METHOD PRIVATE Test_EStopRequestSwitchesOutputsOffAndBlocksRestart
TcUnit.TEST(__POUNAME());
// arrange: running
group_3(Run := TRUE);
fb_3(Restart := FALSE, EStopIn1 := TRUE, EStopIn2 := TRUE);
group_3(Run := TRUE);
fb_3(Restart := TRUE, EStopIn1 := TRUE, EStopIn2 := TRUE);
group_3(Run := TRUE);
fb_3(Restart := FALSE, EStopIn1 := TRUE, EStopIn2 := TRUE);
// act: press the e-stop
group_3(Run := TRUE);
fb_3(Restart := FALSE, EStopIn1 := FALSE, EStopIn2 := FALSE);
// assert
AssertEquals_BOOL(Expected := FALSE, Actual := fb_3.EStopOut, Message := 'EStopOut off');
AssertEquals_BOOL(Expected := FALSE, Actual := fb_3.EStopDelOut, Message := 'EStopDelOut off without delay time');
AssertEquals_BYTE(Expected := TO_BYTE(E_SafeFbState.Safe), Actual := fb_3.State, Message := 'state SAFE');
// act: restart while still pressed
group_3(Run := TRUE);
fb_3(Restart := TRUE, EStopIn1 := FALSE, EStopIn2 := FALSE);
group_3(Run := TRUE);
fb_3(Restart := FALSE, EStopIn1 := FALSE, EStopIn2 := FALSE);
AssertEquals_BOOL(Expected := FALSE, Actual := fb_3.EStopOut, Message := 'restart ignored while the e-stop is pressed');
TEST_FINISHED_NAMED(__POUNAME());
END_METHOD

METHOD PRIVATE Test_MakeContactInputRequestsSafeStateOnOne
TcUnit.TEST(__POUNAME());
// arrange: single channel make contact, released (0), restarted
group_4(Run := TRUE);
fb_4(Restart := FALSE, EStopIn1 := FALSE);
group_4(Run := TRUE);
fb_4(Restart := TRUE, EStopIn1 := FALSE);
group_4(Run := TRUE);
fb_4(Restart := FALSE, EStopIn1 := FALSE);
AssertEquals_BYTE(Expected := TO_BYTE(E_SafeFbState.Run), Actual := fb_4.State, Message := 'running with make contact released');
// act
group_4(Run := TRUE);
fb_4(Restart := FALSE, EStopIn1 := TRUE);
// assert
AssertEquals_BYTE(Expected := TO_BYTE(E_SafeFbState.Safe), Actual := fb_4.State, Message := 'make contact at 1 requests the safe state');
TEST_FINISHED_NAMED(__POUNAME());
END_METHOD

METHOD PRIVATE Test_OutputsOffWhenStopped
TcUnit.TEST(__POUNAME());
// act
group_1(Run := FALSE);
fb_1(EStopIn1 := TRUE);
// assert
AssertEquals_BOOL(Expected := FALSE, Actual := fb_1.EStopOut, Message := 'no output while the group is stopped');
AssertEquals_BYTE(Expected := TO_BYTE(E_SafeFbState.Stop), Actual := fb_1.State, Message := 'state STOP');
TEST_FINISHED_NAMED(__POUNAME());
END_METHOD

METHOD PRIVATE Test_ResetTimeOverSixtySecondsIsRefused
TcUnit.TEST(__POUNAME());
// arrange / act: Edm2ResetTime is 60010 ms, which the Safety Editor refuses
group_9(Run := TRUE);
fb_9(EDM2 := TRUE, EStopIn1 := TRUE);
group_9(Run := TRUE);
fb_9(EDM2 := TRUE, EStopIn1 := TRUE);
// assert
AssertEquals_BOOL(Expected := TRUE, Actual := fb_9.Error, Message := 'configuration error reported');
AssertEquals_BYTE(Expected := TO_BYTE(E_SafeFbState.Error), Actual := fb_9.State, Message := 'state ERROR');
AssertEquals_WORD(Expected := WORD#16#8000, Actual := fb_9.Diag, Message := 'diag bit 15 configuration refused');
AssertEquals_BOOL(Expected := FALSE, Actual := fb_9.EStopOut, Message := 'EStopOut stays at its safe value');
AssertEquals_BOOL(Expected := TRUE, Actual := group_9.FbErr, Message := 'the group sees an FB error');
// act: ErrAck 0 -> 1 -> 0 does not clear a configuration error
group_9(Run := TRUE, ErrAck := TRUE);
fb_9(EDM2 := TRUE, EStopIn1 := TRUE);
group_9(Run := TRUE, ErrAck := TRUE);
fb_9(EDM2 := TRUE, EStopIn1 := TRUE);
group_9(Run := TRUE, ErrAck := FALSE);
fb_9(EDM2 := TRUE, EStopIn1 := TRUE);
AssertEquals_BOOL(Expected := TRUE, Actual := fb_9.Error, Message := 'error not acknowledged');
AssertEquals_WORD(Expected := WORD#16#8000, Actual := fb_9.Diag, Message := 'diag bit 15 kept');
TEST_FINISHED_NAMED(__POUNAME());
END_METHOD

METHOD PRIVATE Test_RestartHeldBeforeEStopGivesEdmError
TcUnit.TEST(__POUNAME());
// arrange: running with EDM feedback (contactors pulled in -> EDM1 = 0)
group_6(Run := TRUE);
fb_6(Restart := FALSE, EDM1 := TRUE, EStopIn1 := TRUE);
group_6(Run := TRUE);
fb_6(Restart := TRUE, EDM1 := TRUE, EStopIn1 := TRUE);
group_6(Run := TRUE);
fb_6(Restart := FALSE, EDM1 := TRUE, EStopIn1 := TRUE);
group_6(Run := TRUE);
fb_6(Restart := FALSE, EDM1 := FALSE, EStopIn1 := TRUE);
// act: restart held, then e-stop pressed before the contactors drop out
group_6(Run := TRUE);
fb_6(Restart := TRUE, EDM1 := FALSE, EStopIn1 := FALSE);
// assert
AssertEquals_BOOL(Expected := TRUE, Actual := fb_6.Error, Message := 'immediate EDM check with restart held (sample 3)');
TEST_FINISHED_NAMED(__POUNAME());
END_METHOD

METHOD PRIVATE Test_StartupRequiresRestartSequence
TcUnit.TEST(__POUNAME());
// act: two channel e-stop released, no restart yet
group_2(Run := TRUE);
fb_2(Restart := FALSE, EStopIn1 := TRUE, EStopIn2 := TRUE);
group_2(Run := TRUE);
fb_2(Restart := FALSE, EStopIn1 := TRUE, EStopIn2 := TRUE);
// assert
AssertEquals_BOOL(Expected := FALSE, Actual := fb_2.EStopOut, Message := 'no output before restart');
AssertEquals_BYTE(Expected := TO_BYTE(E_SafeFbState.Safe), Actual := fb_2.State, Message := 'state SAFE waiting for restart');
group_2(Run := TRUE);
fb_2(Restart := TRUE, EStopIn1 := TRUE, EStopIn2 := TRUE);
AssertEquals_BYTE(Expected := TO_BYTE(E_SafeFbState.Start), Actual := fb_2.State, Message := 'state START while restart held');
AssertEquals_BOOL(Expected := FALSE, Actual := fb_2.EStopOut, Message := 'no output while restart held');
group_2(Run := TRUE);
fb_2(Restart := FALSE, EStopIn1 := TRUE, EStopIn2 := TRUE);
AssertEquals_BYTE(Expected := TO_BYTE(E_SafeFbState.Run), Actual := fb_2.State, Message := 'state RUN after falling edge');
AssertEquals_BOOL(Expected := TRUE, Actual := fb_2.EStopOut, Message := 'EStopOut on');
AssertEquals_BOOL(Expected := TRUE, Actual := fb_2.EStopDelOut, Message := 'EStopDelOut on');
TEST_FINISHED_NAMED(__POUNAME());
END_METHOD

END_FUNCTION_BLOCK

// Tests/T_SafeMon_Tests
FUNCTION_BLOCK T_SafeMon_Tests EXTENDS TcUnit.FB_TestSuite
VAR
    // Test_AutomaticRestartWhenGuardClosed
    group_1 : T_SafeGroup;
    fb_1 : T_SafeMon(group := group_1);
    // Test_SecureInputBypassesGuard
    group_2 : T_SafeGroup;
    fb_2 : T_SafeMon(group := group_2);
    // Test_ManualFunctionTestRequiresGuardOpenedOnce
    group_3 : T_SafeGroup;
    fb_3 : T_SafeMon(group := group_3) := (Parameters := (ManualFunctionTest := TRUE));
    // Test_EdmFaultWithoutManualRestartStaysSafe
    group_4 : T_SafeGroup;
    fb_4 : T_SafeMon(group := group_4);
    // Test_NoMonInConnectedIsRefused
    group_5 : T_SafeGroup;
    fb_5 : T_SafeMon(group := group_5);
    // Test_ResetTimeNotMultipleOfTenIsRefused
    group_6 : T_SafeGroup;
    fb_6 : T_SafeMon(group := group_6) := (Parameters := (Edm1ResetTime := T#15MS));
END_VAR

Test_AutomaticRestartWhenGuardClosed();
Test_SecureInputBypassesGuard();
Test_ManualFunctionTestRequiresGuardOpenedOnce();
Test_EdmFaultWithoutManualRestartStaysSafe();
Test_NoMonInConnectedIsRefused();
Test_ResetTimeNotMultipleOfTenIsRefused();

METHOD PRIVATE Test_AutomaticRestartWhenGuardClosed
TcUnit.TEST(__POUNAME());
// act: Restart not connected -> automatic restart; guard open
group_1(Run := TRUE);
fb_1(MonIn1 := FALSE);
group_1(Run := TRUE);
fb_1(MonIn1 := FALSE);
// assert
AssertEquals_BOOL(Expected := FALSE, Actual := fb_1.MonOut, Message := 'output off with guard open');
group_1(Run := TRUE);
fb_1(MonIn1 := TRUE);
AssertEquals_BOOL(Expected := TRUE, Actual := fb_1.MonOut, Message := 'automatic restart with guard closed');
AssertEquals_BYTE(Expected := TO_BYTE(E_SafeMonState.Run), Actual := fb_1.State, Message := 'state RUN');
TEST_FINISHED_NAMED(__POUNAME());
END_METHOD

METHOD PRIVATE Test_EdmFaultWithoutManualRestartStaysSafe
TcUnit.TEST(__POUNAME());
// act: EDM1 connected and FALSE, no Restart connected
group_4(Run := TRUE);
fb_4(EDM1 := FALSE, MonIn1 := TRUE);
group_4(Run := TRUE);
fb_4(EDM1 := FALSE, MonIn1 := TRUE);
// assert
AssertEquals_BOOL(Expected := FALSE, Actual := fb_4.Error, Message := 'no EDM error without manual restart');
AssertEquals_BYTE(Expected := TO_BYTE(E_SafeMonState.Safe), Actual := fb_4.State, Message := 'FB remains SAFE');
TEST_FINISHED_NAMED(__POUNAME());
END_METHOD

METHOD PRIVATE Test_ManualFunctionTestRequiresGuardOpenedOnce
TcUnit.TEST(__POUNAME());
// arrange: Restart connected (manual restart), guard closed from the start
group_3(Run := TRUE);
fb_3(Restart := FALSE, MonIn1 := TRUE);
AssertEquals_BYTE(Expected := TO_BYTE(E_SafeMonState.FuncTest), Actual := fb_3.State, Message := 'state FUNCTEST after start');
// act: restart without testing the guard
group_3(Run := TRUE);
fb_3(Restart := TRUE, MonIn1 := TRUE);
group_3(Run := TRUE);
fb_3(Restart := FALSE, MonIn1 := TRUE);
AssertEquals_BOOL(Expected := FALSE, Actual := fb_3.MonOut, Message := 'restart ignored before the function test');
// act: open and close the guard, then restart
group_3(Run := TRUE);
fb_3(Restart := FALSE, MonIn1 := FALSE);
group_3(Run := TRUE);
fb_3(Restart := FALSE, MonIn1 := TRUE);
group_3(Run := TRUE);
fb_3(Restart := TRUE, MonIn1 := TRUE);
group_3(Run := TRUE);
fb_3(Restart := FALSE, MonIn1 := TRUE);
AssertEquals_BOOL(Expected := TRUE, Actual := fb_3.MonOut, Message := 'output on after function test and restart');
TEST_FINISHED_NAMED(__POUNAME());
END_METHOD

METHOD PRIVATE Test_NoMonInConnectedIsRefused
TcUnit.TEST(__POUNAME());
// arrange / act: only the Secure pair is connected, which the Safety Editor refuses
group_5(Run := TRUE);
fb_5(Secure1 := TRUE);
group_5(Run := TRUE);
fb_5(Secure1 := TRUE);
// assert
AssertEquals_BOOL(Expected := TRUE, Actual := fb_5.Error, Message := 'configuration error reported');
AssertEquals_BYTE(Expected := TO_BYTE(E_SafeFbState.Error), Actual := fb_5.State, Message := 'state ERROR');
AssertEquals_WORD(Expected := WORD#16#8000, Actual := fb_5.Diag, Message := 'diag bit 15 configuration refused');
AssertEquals_BOOL(Expected := FALSE, Actual := fb_5.MonOut, Message := 'MonOut stays at its safe value');
AssertEquals_BOOL(Expected := TRUE, Actual := group_5.FbErr, Message := 'the group sees an FB error');
// act: ErrAck 0 -> 1 -> 0 does not clear a configuration error
group_5(Run := TRUE, ErrAck := TRUE);
fb_5(Secure1 := TRUE);
group_5(Run := TRUE, ErrAck := TRUE);
fb_5(Secure1 := TRUE);
group_5(Run := TRUE, ErrAck := FALSE);
fb_5(Secure1 := TRUE);
AssertEquals_BOOL(Expected := TRUE, Actual := fb_5.Error, Message := 'error not acknowledged');
AssertEquals_WORD(Expected := WORD#16#8000, Actual := fb_5.Diag, Message := 'diag bit 15 kept');
TEST_FINISHED_NAMED(__POUNAME());
END_METHOD

METHOD PRIVATE Test_ResetTimeNotMultipleOfTenIsRefused
TcUnit.TEST(__POUNAME());
// arrange / act: Edm1ResetTime is 15 ms, which the Safety Editor refuses
group_6(Run := TRUE);
fb_6(EDM1 := TRUE, MonIn1 := TRUE);
group_6(Run := TRUE);
fb_6(EDM1 := TRUE, MonIn1 := TRUE);
// assert
AssertEquals_BOOL(Expected := TRUE, Actual := fb_6.Error, Message := 'configuration error reported');
AssertEquals_BYTE(Expected := TO_BYTE(E_SafeFbState.Error), Actual := fb_6.State, Message := 'state ERROR');
AssertEquals_WORD(Expected := WORD#16#8000, Actual := fb_6.Diag, Message := 'diag bit 15 configuration refused');
AssertEquals_BOOL(Expected := FALSE, Actual := fb_6.MonOut, Message := 'MonOut stays at its safe value');
AssertEquals_BOOL(Expected := TRUE, Actual := group_6.FbErr, Message := 'the group sees an FB error');
// act: ErrAck 0 -> 1 -> 0 does not clear a configuration error
group_6(Run := TRUE, ErrAck := TRUE);
fb_6(EDM1 := TRUE, MonIn1 := TRUE);
group_6(Run := TRUE, ErrAck := TRUE);
fb_6(EDM1 := TRUE, MonIn1 := TRUE);
group_6(Run := TRUE, ErrAck := FALSE);
fb_6(EDM1 := TRUE, MonIn1 := TRUE);
AssertEquals_BOOL(Expected := TRUE, Actual := fb_6.Error, Message := 'error not acknowledged');
AssertEquals_WORD(Expected := WORD#16#8000, Actual := fb_6.Diag, Message := 'diag bit 15 kept');
TEST_FINISHED_NAMED(__POUNAME());
END_METHOD

METHOD PRIVATE Test_SecureInputBypassesGuard
TcUnit.TEST(__POUNAME());
// act: guard open, bypass active
group_2(Run := TRUE);
fb_2(MonIn1 := FALSE, Secure1 := TRUE);
group_2(Run := TRUE);
fb_2(MonIn1 := FALSE, Secure1 := TRUE);
// assert
AssertEquals_BOOL(Expected := TRUE, Actual := fb_2.MonOut, Message := 'guard ignored while Secure is 1');
group_2(Run := TRUE);
fb_2(MonIn1 := FALSE, Secure1 := FALSE);
AssertEquals_BOOL(Expected := FALSE, Actual := fb_2.MonOut, Message := 'guard monitored again when Secure is 0');
TEST_FINISHED_NAMED(__POUNAME());
END_METHOD

END_FUNCTION_BLOCK

// Tests/T_SafeTwoHand_Tests
FUNCTION_BLOCK T_SafeTwoHand_Tests EXTENDS TcUnit.FB_TestSuite
VAR
    // Test_BothHandsGiveOutputAndReleaseNeedsBothOff
    group_1 : T_SafeGroup;
    fb_1 : T_SafeTwoHand(group := group_1);
    // Test_SecondHandWithoutFirstGivesTwoHandError
    group_2 : T_SafeGroup;
    fb_2 : T_SafeTwoHand(group := group_2);
    // Test_HandDiscrepancyTimeout
    group_3 : T_SafeGroup;
    // SafeInputsAfterDiscError TRUE (not the default) so the error waits for both hands released (diag bit 10)
    fb_3 : T_SafeTwoHand(group := group_3) := (Parameters := (HandDiscrepancyTime := T#100MS, SafeInputsAfterDiscError := TRUE));
    state_3 : INT := 10;
    waitTimer_3 : TON;
END_VAR

Test_BothHandsGiveOutputAndReleaseNeedsBothOff();
Test_SecondHandWithoutFirstGivesTwoHandError();
Test_HandDiscrepancyTimeout();

METHOD PRIVATE Test_BothHandsGiveOutputAndReleaseNeedsBothOff
TcUnit.TEST(__POUNAME());
// arrange: single channel per hand
group_1(Run := TRUE);
fb_1(Twohand1 := FALSE, Twohand3 := FALSE);
// act
group_1(Run := TRUE);
fb_1(Twohand1 := TRUE, Twohand3 := FALSE);
AssertEquals_BYTE(Expected := TO_BYTE(E_SafeTwoHandState.OneButton), Actual := fb_1.State, Message := 'state 1BUTTON');
group_1(Run := TRUE);
fb_1(Twohand1 := TRUE, Twohand3 := TRUE);
// assert
AssertEquals_BOOL(Expected := TRUE, Actual := fb_1.TwoHandOut, Message := 'output on with both hands');
group_1(Run := TRUE);
fb_1(Twohand1 := FALSE, Twohand3 := TRUE);
AssertEquals_BOOL(Expected := FALSE, Actual := fb_1.TwoHandOut, Message := 'output off when one hand released');
AssertEquals_BYTE(Expected := TO_BYTE(E_SafeTwoHandState.Release), Actual := fb_1.State, Message := 'state RELEASE');
group_1(Run := TRUE);
fb_1(Twohand1 := TRUE, Twohand3 := TRUE);
AssertEquals_BOOL(Expected := FALSE, Actual := fb_1.TwoHandOut, Message := 'no re-trigger until both hands released');
TEST_FINISHED_NAMED(__POUNAME());
END_METHOD

METHOD PRIVATE Test_HandDiscrepancyTimeout
TcUnit.TEST(__POUNAME());
waitTimer_3();

CASE state_3 OF
    10:
        group_3(Run := TRUE);
        fb_3(Twohand1 := FALSE, Twohand3 := FALSE);
        state_3 := 20;
        waitTimer_3(IN := TRUE, PT := T#250MS);
    20:
        // act: only one hand for longer than the discrepancy time
        group_3(Run := TRUE);
        fb_3(Twohand1 := TRUE, Twohand3 := FALSE);

        IF NOT waitTimer_3.Q THEN
            RETURN;
        END_IF

        waitTimer_3(IN := FALSE);
        // assert
        AssertEquals_BOOL(Expected := TRUE, Actual := fb_3.Error, Message := 'discrepancy error between hands');
        AssertEquals_WORD(Expected := WORD#16#0404, Actual := fb_3.Diag, Message := 'diag bits 2 and 10');
        TEST_FINISHED_NAMED(__POUNAME());
        state_3 := 10;
END_CASE
END_METHOD

METHOD PRIVATE Test_SecondHandWithoutFirstGivesTwoHandError
TcUnit.TEST(__POUNAME());
// arrange
group_2(Run := TRUE);
fb_2(Twohand1 := FALSE, Twohand3 := FALSE);
group_2(Run := TRUE);
fb_2(Twohand1 := TRUE, Twohand3 := FALSE);
// act: first hand lost as the second is actuated
group_2(Run := TRUE);
fb_2(Twohand1 := FALSE, Twohand3 := TRUE);
// assert
AssertEquals_BOOL(Expected := TRUE, Actual := fb_2.Error, Message := 'two-hand error');
AssertEquals_WORD(Expected := WORD#64, Actual := fb_2.Diag, Message := 'diag bit 6');
TEST_FINISHED_NAMED(__POUNAME());
END_METHOD

END_FUNCTION_BLOCK

// Tests/T_SafeMuting_Tests
FUNCTION_BLOCK T_SafeMuting_Tests EXTENDS TcUnit.FB_TestSuite
VAR
    // Test_OssdBlockedWithoutMutingGivesSafe
    group_1 : T_SafeGroup;
    fb_1 : T_SafeMuting(group := group_1);
    // Test_SequentialMutingKeepsOutputOn
    group_2 : T_SafeGroup;
    fb_2 : T_SafeMuting(group := group_2) := (Parameters := (SequentialInputs := TRUE));
    // Test_SequenceViolationGivesError
    group_3 : T_SafeGroup;
    fb_3 : T_SafeMuting(group := group_3) := (Parameters := (SequentialInputs := TRUE));
    // Test_TwoSensorParallelSequence
    group_4 : T_SafeGroup;
    fb_4 : T_SafeMuting(group := group_4);
    // Test_ResetTimeNotMultipleOfTenIsRefused
    group_5 : T_SafeGroup;
    fb_5 : T_SafeMuting(group := group_5) := (Parameters := (Edm1ResetTime := T#25MS));
END_VAR

Test_OssdBlockedWithoutMutingGivesSafe();
Test_SequentialMutingKeepsOutputOn();
Test_SequenceViolationGivesError();
Test_TwoSensorParallelSequence();
Test_ResetTimeNotMultipleOfTenIsRefused();

METHOD PRIVATE Test_OssdBlockedWithoutMutingGivesSafe
TcUnit.TEST(__POUNAME());
// arrange: only the protective device connected
group_1(Run := TRUE);
fb_1(OSSDIn1 := TRUE);
group_1(Run := TRUE);
fb_1(OSSDIn1 := TRUE);
AssertEquals_BOOL(Expected := TRUE, Actual := fb_1.MuteOut, Message := 'output on with clear protective device');
// act
group_1(Run := TRUE);
fb_1(OSSDIn1 := FALSE);
// assert
AssertEquals_BOOL(Expected := FALSE, Actual := fb_1.MuteOut, Message := 'output off when interrupted');
AssertEquals_BYTE(Expected := TO_BYTE(E_SafeMutingState.Safe), Actual := fb_1.State, Message := 'state SAFE');
group_1(Run := TRUE);
fb_1(OSSDIn1 := TRUE);
AssertEquals_BOOL(Expected := TRUE, Actual := fb_1.MuteOut, Message := 'automatic restart when clear again');
TEST_FINISHED_NAMED(__POUNAME());
END_METHOD

METHOD PRIVATE Test_ResetTimeNotMultipleOfTenIsRefused
TcUnit.TEST(__POUNAME());
// arrange / act: Edm1ResetTime is 25 ms, which the Safety Editor refuses
group_5(Run := TRUE);
fb_5(EDM1 := TRUE, OSSDIn1 := TRUE);
group_5(Run := TRUE);
fb_5(EDM1 := TRUE, OSSDIn1 := TRUE);
// assert
AssertEquals_BOOL(Expected := TRUE, Actual := fb_5.Error, Message := 'configuration error reported');
AssertEquals_BYTE(Expected := TO_BYTE(E_SafeFbState.Error), Actual := fb_5.State, Message := 'state ERROR');
AssertEquals_WORD(Expected := WORD#16#8000, Actual := fb_5.Diag, Message := 'diag bit 15 configuration refused');
AssertEquals_BOOL(Expected := FALSE, Actual := fb_5.MuteOut, Message := 'MuteOut stays at its safe value');
AssertEquals_BOOL(Expected := TRUE, Actual := group_5.FbErr, Message := 'the group sees an FB error');
// act: ErrAck 0 -> 1 -> 0 does not clear a configuration error
group_5(Run := TRUE, ErrAck := TRUE);
fb_5(EDM1 := TRUE, OSSDIn1 := TRUE);
group_5(Run := TRUE, ErrAck := TRUE);
fb_5(EDM1 := TRUE, OSSDIn1 := TRUE);
group_5(Run := TRUE, ErrAck := FALSE);
fb_5(EDM1 := TRUE, OSSDIn1 := TRUE);
AssertEquals_BOOL(Expected := TRUE, Actual := fb_5.Error, Message := 'error not acknowledged');
AssertEquals_WORD(Expected := WORD#16#8000, Actual := fb_5.Diag, Message := 'diag bit 15 kept');
TEST_FINISHED_NAMED(__POUNAME());
END_METHOD

METHOD PRIVATE Test_SequenceViolationGivesError
TcUnit.TEST(__POUNAME());
// arrange
group_3(Run := TRUE);
fb_3(
    MutingEnable := TRUE,
    MutingIn1 := FALSE,
    MutingIn2 := FALSE,
    MutingIn3 := FALSE,
    MutingIn4 := FALSE,
    OSSDIn1 := TRUE
);

group_3(Run := TRUE);
fb_3(
    MutingEnable := TRUE,
    MutingIn1 := FALSE,
    MutingIn2 := FALSE,
    MutingIn3 := FALSE,
    MutingIn4 := FALSE,
    OSSDIn1 := TRUE
);

group_3(Run := TRUE);
fb_3(
    MutingEnable := TRUE,
    MutingIn1 := TRUE,
    MutingIn2 := FALSE,
    MutingIn3 := FALSE,
    MutingIn4 := FALSE,
    OSSDIn1 := TRUE
);

// act: OSSD blocked before the second sensor
group_3(Run := TRUE);
fb_3(
    MutingEnable := TRUE,
    MutingIn1 := TRUE,
    MutingIn2 := FALSE,
    MutingIn3 := FALSE,
    MutingIn4 := FALSE,
    OSSDIn1 := FALSE
);

// assert
AssertEquals_BOOL(Expected := TRUE, Actual := fb_3.Error, Message := 'sequence violation');
AssertEquals_WORD(Expected := WORD#64, Actual := fb_3.Diag, Message := 'diag bit 6');
AssertEquals_BOOL(Expected := FALSE, Actual := fb_3.MuteOut, Message := 'output off');
TEST_FINISHED_NAMED(__POUNAME());
END_METHOD

METHOD PRIVATE Test_SequentialMutingKeepsOutputOn
TcUnit.TEST(__POUNAME());
// arrange: four single-channel sensors, running
group_2(Run := TRUE);
fb_2(
    MutingEnable := TRUE,
    MutingIn1 := FALSE,
    MutingIn2 := FALSE,
    MutingIn3 := FALSE,
    MutingIn4 := FALSE,
    OSSDIn1 := TRUE
);

group_2(Run := TRUE);
fb_2(
    MutingEnable := TRUE,
    MutingIn1 := FALSE,
    MutingIn2 := FALSE,
    MutingIn3 := FALSE,
    MutingIn4 := FALSE,
    OSSDIn1 := TRUE
);

// act: M1, M2, OSSD blocked, M3, M1 off, M4, M2 off, OSSD clear, M3 off, M4 off
group_2(Run := TRUE);
fb_2(
    MutingEnable := TRUE,
    MutingIn1 := TRUE,
    MutingIn2 := FALSE,
    MutingIn3 := FALSE,
    MutingIn4 := FALSE,
    OSSDIn1 := TRUE
);

AssertEquals_BYTE(Expected := TO_BYTE(E_SafeMutingState.Muting1), Actual := fb_2.State, Message := 'MUTING1');
AssertEquals_BOOL(Expected := TRUE, Actual := fb_2.MutingActive, Message := 'muting active');
group_2(Run := TRUE);
fb_2(
    MutingEnable := TRUE,
    MutingIn1 := TRUE,
    MutingIn2 := TRUE,
    MutingIn3 := FALSE,
    MutingIn4 := FALSE,
    OSSDIn1 := TRUE
);

group_2(Run := TRUE);
fb_2(
    MutingEnable := TRUE,
    MutingIn1 := TRUE,
    MutingIn2 := TRUE,
    MutingIn3 := FALSE,
    MutingIn4 := FALSE,
    OSSDIn1 := FALSE
);

AssertEquals_BYTE(Expected := TO_BYTE(E_SafeMutingState.Muting3), Actual := fb_2.State, Message := 'MUTING3');
AssertEquals_BOOL(Expected := TRUE, Actual := fb_2.MuteOut, Message := 'output stays on while muted');
group_2(Run := TRUE);
fb_2(
    MutingEnable := TRUE,
    MutingIn1 := TRUE,
    MutingIn2 := TRUE,
    MutingIn3 := TRUE,
    MutingIn4 := FALSE,
    OSSDIn1 := FALSE
);

group_2(Run := TRUE);
fb_2(
    MutingEnable := TRUE,
    MutingIn1 := FALSE,
    MutingIn2 := TRUE,
    MutingIn3 := TRUE,
    MutingIn4 := FALSE,
    OSSDIn1 := FALSE
);

group_2(Run := TRUE);
fb_2(
    MutingEnable := TRUE,
    MutingIn1 := FALSE,
    MutingIn2 := TRUE,
    MutingIn3 := TRUE,
    MutingIn4 := TRUE,
    OSSDIn1 := FALSE
);

group_2(Run := TRUE);
fb_2(
    MutingEnable := TRUE,
    MutingIn1 := FALSE,
    MutingIn2 := FALSE,
    MutingIn3 := TRUE,
    MutingIn4 := TRUE,
    OSSDIn1 := FALSE
);

group_2(Run := TRUE);
fb_2(
    MutingEnable := TRUE,
    MutingIn1 := FALSE,
    MutingIn2 := FALSE,
    MutingIn3 := TRUE,
    MutingIn4 := TRUE,
    OSSDIn1 := TRUE
);

AssertEquals_BYTE(Expected := TO_BYTE(E_SafeMutingState.Muting8), Actual := fb_2.State, Message := 'MUTING8');
group_2(Run := TRUE);
fb_2(
    MutingEnable := TRUE,
    MutingIn1 := FALSE,
    MutingIn2 := FALSE,
    MutingIn3 := FALSE,
    MutingIn4 := TRUE,
    OSSDIn1 := TRUE
);

group_2(Run := TRUE);
fb_2(
    MutingEnable := TRUE,
    MutingIn1 := FALSE,
    MutingIn2 := FALSE,
    MutingIn3 := FALSE,
    MutingIn4 := FALSE,
    OSSDIn1 := TRUE
);

// assert
AssertEquals_BYTE(Expected := TO_BYTE(E_SafeMutingState.Run), Actual := fb_2.State, Message := 'RUN after the sequence');
AssertEquals_BOOL(Expected := FALSE, Actual := fb_2.MutingActive, Message := 'muting no longer active');
AssertEquals_BOOL(Expected := FALSE, Actual := fb_2.Error, Message := 'no error');
TEST_FINISHED_NAMED(__POUNAME());
END_METHOD

METHOD PRIVATE Test_TwoSensorParallelSequence
TcUnit.TEST(__POUNAME());
// arrange: two two-channel sensors (parallel inputs), running
group_4(Run := TRUE);
fb_4(
    MutingEnable := TRUE,
    MutingIn1 := FALSE,
    MutingIn2 := FALSE,
    MutingIn3 := FALSE,
    MutingIn4 := FALSE,
    OSSDIn1 := TRUE
);

group_4(Run := TRUE);
fb_4(
    MutingEnable := TRUE,
    MutingIn1 := FALSE,
    MutingIn2 := FALSE,
    MutingIn3 := FALSE,
    MutingIn4 := FALSE,
    OSSDIn1 := TRUE
);

// act: S1, S2, OSSD blocked, S1 off, OSSD clear, S2 off
group_4(Run := TRUE);
fb_4(
    MutingEnable := TRUE,
    MutingIn1 := TRUE,
    MutingIn2 := TRUE,
    MutingIn3 := FALSE,
    MutingIn4 := FALSE,
    OSSDIn1 := TRUE
);

group_4(Run := TRUE);
fb_4(
    MutingEnable := TRUE,
    MutingIn1 := TRUE,
    MutingIn2 := TRUE,
    MutingIn3 := TRUE,
    MutingIn4 := TRUE,
    OSSDIn1 := TRUE
);

group_4(Run := TRUE);
fb_4(
    MutingEnable := TRUE,
    MutingIn1 := TRUE,
    MutingIn2 := TRUE,
    MutingIn3 := TRUE,
    MutingIn4 := TRUE,
    OSSDIn1 := FALSE
);

AssertEquals_BOOL(Expected := TRUE, Actual := fb_4.MuteOut, Message := 'output stays on while muted');
group_4(Run := TRUE);
fb_4(
    MutingEnable := TRUE,
    MutingIn1 := FALSE,
    MutingIn2 := FALSE,
    MutingIn3 := TRUE,
    MutingIn4 := TRUE,
    OSSDIn1 := FALSE
);

group_4(Run := TRUE);
fb_4(
    MutingEnable := TRUE,
    MutingIn1 := FALSE,
    MutingIn2 := FALSE,
    MutingIn3 := TRUE,
    MutingIn4 := TRUE,
    OSSDIn1 := TRUE
);

group_4(Run := TRUE);
fb_4(
    MutingEnable := TRUE,
    MutingIn1 := FALSE,
    MutingIn2 := FALSE,
    MutingIn3 := FALSE,
    MutingIn4 := FALSE,
    OSSDIn1 := TRUE
);

// assert
AssertEquals_BYTE(Expected := TO_BYTE(E_SafeMutingState.Run), Actual := fb_4.State, Message := 'RUN after the sequence');
AssertEquals_BOOL(Expected := FALSE, Actual := fb_4.Error, Message := 'no error');
TEST_FINISHED_NAMED(__POUNAME());
END_METHOD

END_FUNCTION_BLOCK

// Tests/T_SafeConnection_Tests
FUNCTION_BLOCK T_SafeConnection_Tests EXTENDS TcUnit.FB_TestSuite
VAR
    // Test_StartsUpToDataWhenGroupRuns
    group_1 : T_SafeGroup;
    conn_1 : T_SafeConnection(group := group_1);
    i_1 : INT;
    // Test_ComErrorClearedByAcknowledge
    group_2 : T_SafeGroup;
    conn_2 : T_SafeConnection(group := group_2);
    i_2 : INT;
END_VAR

Test_StartsUpToDataWhenGroupRuns();
Test_ComErrorClearedByAcknowledge();

METHOD PRIVATE Test_ComErrorClearedByAcknowledge
VAR
    diag : BYTE;
END_VAR
TcUnit.TEST(__POUNAME());

// arrange
FOR i_2 := 1 TO 5 DO
    group_2(Run := TRUE, ErrAck := FALSE);
    conn_2(InjectComError := FALSE, StartupTime := T#0S);
END_FOR

// act
group_2(Run := TRUE, ErrAck := FALSE);
conn_2(InjectComError := TRUE, StartupTime := T#0S);
// assert
AssertEquals_BOOL(Expected := TRUE, Actual := conn_2.ComError, Message := 'com error');
AssertEquals_BOOL(Expected := FALSE, Actual := conn_2.InDataState, Message := 'dropped out of Data');
diag := conn_2.Diag AND 16#0F;
AssertEquals_BYTE(Expected := BYTE#5, Actual := diag, Message := 'diag code watchdog');
group_2(Run := TRUE, ErrAck := FALSE);
conn_2(InjectComError := FALSE, StartupTime := T#0S);
AssertEquals_BYTE(Expected := TO_BYTE(E_SafeGroupState.Error), Actual := group_2.State, Message := 'group ERROR');
group_2(Run := TRUE, ErrAck := TRUE);
conn_2(InjectComError := FALSE, StartupTime := T#0S);

FOR i_2 := 1 TO 5 DO
    group_2(Run := TRUE, ErrAck := FALSE);
    conn_2(InjectComError := FALSE, StartupTime := T#0S);
END_FOR

AssertEquals_BOOL(Expected := FALSE, Actual := conn_2.ComError, Message := 'error cleared');
AssertEquals_BOOL(Expected := TRUE, Actual := conn_2.InDataState, Message := 'restarted to Data');
TEST_FINISHED_NAMED(__POUNAME());
END_METHOD

METHOD PRIVATE Test_StartsUpToDataWhenGroupRuns
TcUnit.TEST(__POUNAME());
// act
group_1(Run := FALSE);
conn_1(StartupTime := T#0S);
AssertEquals_BOOL(Expected := TRUE, Actual := conn_1.InStartup, Message := 'in startup before the group runs');

FOR i_1 := 1 TO 5 DO
    group_1(Run := TRUE);
    conn_1(StartupTime := T#0S);
END_FOR

// assert
AssertEquals_BOOL(Expected := TRUE, Actual := conn_1.InDataState, Message := 'Data state reached');
AssertEquals_BOOL(Expected := FALSE, Actual := conn_1.InStartup, Message := 'no longer in startup');
TEST_FINISHED_NAMED(__POUNAME());
END_METHOD

END_FUNCTION_BLOCK

// Tests/T_SafeInputTerminal8_Tests
FUNCTION_BLOCK T_SafeInputTerminal8_Tests EXTENDS TcUnit.FB_TestSuite
VAR
    // Test_SafeInputsFalseBeforeData
    group_1 : T_SafeGroup;
    terminal_1 : T_SafeInputTerminal8(group := group_1);
    // Test_SafeInputsFollowChannelsInData
    group_2 : T_SafeGroup;
    terminal_2 : T_SafeInputTerminal8(group := group_2);
    i_2 : INT;
    // Test_ComErrorForcesSafeInputsFalse
    group_3 : T_SafeGroup;
    terminal_3 : T_SafeInputTerminal8(group := group_3);
    i_3 : INT;
    // Test_RegistersAsConnection
    group_4 : T_SafeGroup;
    terminal_4 : T_SafeInputTerminal8(group := group_4);
END_VAR

Test_SafeInputsFalseBeforeData();
Test_SafeInputsFollowChannelsInData();
Test_ComErrorForcesSafeInputsFalse();
Test_RegistersAsConnection();

METHOD PRIVATE Test_ComErrorForcesSafeInputsFalse
TcUnit.TEST(__POUNAME());

// arrange: in Data with every channel on
FOR i_3 := 1 TO 5 DO
    group_3(Run := TRUE);
    terminal_3(Channel1 := TRUE, Channel2 := TRUE, Channel3 := TRUE, Channel4 := TRUE,
               Channel5 := TRUE, Channel6 := TRUE, Channel7 := TRUE, Channel8 := TRUE,
               StartupTime := T#0S);
END_FOR
AssertEquals_BOOL(Expected := TRUE, Actual := terminal_3.SafeIn8, Message := 'SafeIn8 on before the error');

// act
group_3(Run := TRUE);
terminal_3(Channel1 := TRUE, Channel2 := TRUE, Channel3 := TRUE, Channel4 := TRUE,
               Channel5 := TRUE, Channel6 := TRUE, Channel7 := TRUE, Channel8 := TRUE,
               InjectComError := TRUE, StartupTime := T#0S);

// assert
AssertEquals_BOOL(Expected := TRUE, Actual := terminal_3.ComError, Message := 'com error');
AssertEquals_BOOL(Expected := FALSE, Actual := terminal_3.SafeIn1, Message := 'SafeIn1 fail-safe on com error');
AssertEquals_BOOL(Expected := FALSE, Actual := terminal_3.SafeIn4, Message := 'SafeIn4 fail-safe on com error');
AssertEquals_BOOL(Expected := FALSE, Actual := terminal_3.SafeIn5, Message := 'SafeIn5 fail-safe on com error');
AssertEquals_BOOL(Expected := FALSE, Actual := terminal_3.SafeIn8, Message := 'SafeIn8 fail-safe on com error');
TEST_FINISHED_NAMED(__POUNAME());
END_METHOD

METHOD PRIVATE Test_RegistersAsConnection
TcUnit.TEST(__POUNAME());

// act
group_4(Run := TRUE);
terminal_4(StartupTime := T#0S);

// assert
AssertEquals_UINT(Expected := 1, Actual := group_4.ConnectionCount, Message := 'one connection registered');
AssertEquals_UINT(Expected := 0, Actual := group_4.FunctionBlockCount, Message := 'no function blocks');
TEST_FINISHED_NAMED(__POUNAME());
END_METHOD

METHOD PRIVATE Test_SafeInputsFalseBeforeData
TcUnit.TEST(__POUNAME());

// arrange: group stopped, so the connection never reaches Data
group_1(Run := FALSE);

// act
terminal_1(Channel1 := TRUE, Channel2 := TRUE, Channel3 := TRUE, Channel4 := TRUE,
           Channel5 := TRUE, Channel6 := TRUE, Channel7 := TRUE, Channel8 := TRUE,
           StartupTime := T#0S);

// assert
AssertEquals_BOOL(Expected := FALSE, Actual := terminal_1.InDataState, Message := 'not in Data');
AssertEquals_BOOL(Expected := FALSE, Actual := terminal_1.SafeIn1, Message := 'SafeIn1 fail-safe');
AssertEquals_BOOL(Expected := FALSE, Actual := terminal_1.SafeIn2, Message := 'SafeIn2 fail-safe');
AssertEquals_BOOL(Expected := FALSE, Actual := terminal_1.SafeIn3, Message := 'SafeIn3 fail-safe');
AssertEquals_BOOL(Expected := FALSE, Actual := terminal_1.SafeIn4, Message := 'SafeIn4 fail-safe');
AssertEquals_BOOL(Expected := FALSE, Actual := terminal_1.SafeIn5, Message := 'SafeIn5 fail-safe');
AssertEquals_BOOL(Expected := FALSE, Actual := terminal_1.SafeIn6, Message := 'SafeIn6 fail-safe');
AssertEquals_BOOL(Expected := FALSE, Actual := terminal_1.SafeIn7, Message := 'SafeIn7 fail-safe');
AssertEquals_BOOL(Expected := FALSE, Actual := terminal_1.SafeIn8, Message := 'SafeIn8 fail-safe');
TEST_FINISHED_NAMED(__POUNAME());
END_METHOD

METHOD PRIVATE Test_SafeInputsFollowChannelsInData
TcUnit.TEST(__POUNAME());

// arrange: run the group until the connection is in Data
FOR i_2 := 1 TO 5 DO
    group_2(Run := TRUE);
    terminal_2(StartupTime := T#0S);
END_FOR
AssertEquals_BOOL(Expected := TRUE, Actual := terminal_2.InDataState, Message := 'Data state reached');

// act: odd channels on, even channels off
group_2(Run := TRUE);
terminal_2(Channel1 := TRUE, Channel2 := FALSE, Channel3 := TRUE, Channel4 := FALSE,
           Channel5 := TRUE, Channel6 := FALSE, Channel7 := TRUE, Channel8 := FALSE,
           StartupTime := T#0S);

// assert
AssertEquals_BOOL(Expected := TRUE, Actual := terminal_2.SafeIn1, Message := 'SafeIn1 follows Channel1');
AssertEquals_BOOL(Expected := FALSE, Actual := terminal_2.SafeIn2, Message := 'SafeIn2 follows Channel2');
AssertEquals_BOOL(Expected := TRUE, Actual := terminal_2.SafeIn3, Message := 'SafeIn3 follows Channel3');
AssertEquals_BOOL(Expected := FALSE, Actual := terminal_2.SafeIn4, Message := 'SafeIn4 follows Channel4');
AssertEquals_BOOL(Expected := TRUE, Actual := terminal_2.SafeIn5, Message := 'SafeIn5 follows Channel5');
AssertEquals_BOOL(Expected := FALSE, Actual := terminal_2.SafeIn6, Message := 'SafeIn6 follows Channel6');
AssertEquals_BOOL(Expected := TRUE, Actual := terminal_2.SafeIn7, Message := 'SafeIn7 follows Channel7');
AssertEquals_BOOL(Expected := FALSE, Actual := terminal_2.SafeIn8, Message := 'SafeIn8 follows Channel8');

// act: invert the pattern
group_2(Run := TRUE);
terminal_2(Channel1 := FALSE, Channel2 := TRUE, Channel3 := FALSE, Channel4 := TRUE,
           Channel5 := FALSE, Channel6 := TRUE, Channel7 := FALSE, Channel8 := TRUE,
           StartupTime := T#0S);

// assert
AssertEquals_BOOL(Expected := FALSE, Actual := terminal_2.SafeIn1, Message := 'SafeIn1 inverted');
AssertEquals_BOOL(Expected := TRUE, Actual := terminal_2.SafeIn2, Message := 'SafeIn2 inverted');
AssertEquals_BOOL(Expected := FALSE, Actual := terminal_2.SafeIn3, Message := 'SafeIn3 inverted');
AssertEquals_BOOL(Expected := TRUE, Actual := terminal_2.SafeIn4, Message := 'SafeIn4 inverted');
AssertEquals_BOOL(Expected := FALSE, Actual := terminal_2.SafeIn5, Message := 'SafeIn5 inverted');
AssertEquals_BOOL(Expected := TRUE, Actual := terminal_2.SafeIn6, Message := 'SafeIn6 inverted');
AssertEquals_BOOL(Expected := FALSE, Actual := terminal_2.SafeIn7, Message := 'SafeIn7 inverted');
AssertEquals_BOOL(Expected := TRUE, Actual := terminal_2.SafeIn8, Message := 'SafeIn8 inverted');
TEST_FINISHED_NAMED(__POUNAME());
END_METHOD

END_FUNCTION_BLOCK

// Tests/T_SafeOutputTerminal2_Tests
FUNCTION_BLOCK T_SafeOutputTerminal2_Tests EXTENDS TcUnit.FB_TestSuite
VAR
    // Test_ChannelsFalseBeforeData
    group_1 : T_SafeGroup;
    terminal_1 : T_SafeOutputTerminal2(group := group_1);
    // Test_ChannelsFollowSafeOutsInData
    group_2 : T_SafeGroup;
    terminal_2 : T_SafeOutputTerminal2(group := group_2);
    i_2 : INT;
    // Test_ComErrorForcesChannelsFalse
    group_3 : T_SafeGroup;
    terminal_3 : T_SafeOutputTerminal2(group := group_3);
    i_3 : INT;
    // Test_RegistersAsConnection
    group_4 : T_SafeGroup;
    terminal_4 : T_SafeOutputTerminal2(group := group_4);
    // Test_GroupNotRunningForcesChannelsFalse
    group_5 : T_SafeGroup;
    terminal_5 : T_SafeOutputTerminal2(group := group_5);
    i_5 : INT;
END_VAR

Test_ChannelsFalseBeforeData();
Test_ChannelsFollowSafeOutsInData();
Test_ComErrorForcesChannelsFalse();
Test_RegistersAsConnection();
Test_GroupNotRunningForcesChannelsFalse();

METHOD PRIVATE Test_ChannelsFalseBeforeData
TcUnit.TEST(__POUNAME());

// arrange: group stopped, so the connection never reaches Data
group_1(Run := FALSE);

// act
terminal_1(SafeOut1 := TRUE, SafeOut2 := TRUE, StartupTime := T#0S);

// assert
AssertEquals_BOOL(Expected := FALSE, Actual := terminal_1.InDataState, Message := 'not in Data');
AssertEquals_BOOL(Expected := FALSE, Actual := terminal_1.Channel1, Message := 'Channel1 fail-safe');
AssertEquals_BOOL(Expected := FALSE, Actual := terminal_1.Channel2, Message := 'Channel2 fail-safe');
TEST_FINISHED_NAMED(__POUNAME());
END_METHOD

METHOD PRIVATE Test_ChannelsFollowSafeOutsInData
TcUnit.TEST(__POUNAME());

// arrange: run the group until the connection is in Data
FOR i_2 := 1 TO 5 DO
    group_2(Run := TRUE);
    terminal_2(StartupTime := T#0S);
END_FOR
AssertEquals_BOOL(Expected := TRUE, Actual := terminal_2.InDataState, Message := 'Data state reached');

// act
group_2(Run := TRUE);
terminal_2(SafeOut1 := TRUE, SafeOut2 := FALSE, StartupTime := T#0S);

// assert
AssertEquals_BOOL(Expected := TRUE, Actual := terminal_2.Channel1, Message := 'Channel1 follows SafeOut1');
AssertEquals_BOOL(Expected := FALSE, Actual := terminal_2.Channel2, Message := 'Channel2 follows SafeOut2');

// act: swap
group_2(Run := TRUE);
terminal_2(SafeOut1 := FALSE, SafeOut2 := TRUE, StartupTime := T#0S);

// assert
AssertEquals_BOOL(Expected := FALSE, Actual := terminal_2.Channel1, Message := 'Channel1 swapped');
AssertEquals_BOOL(Expected := TRUE, Actual := terminal_2.Channel2, Message := 'Channel2 swapped');
TEST_FINISHED_NAMED(__POUNAME());
END_METHOD

METHOD PRIVATE Test_ComErrorForcesChannelsFalse
TcUnit.TEST(__POUNAME());

// arrange: in Data with both outputs on
FOR i_3 := 1 TO 5 DO
    group_3(Run := TRUE);
    terminal_3(SafeOut1 := TRUE, SafeOut2 := TRUE, StartupTime := T#0S);
END_FOR
AssertEquals_BOOL(Expected := TRUE, Actual := terminal_3.Channel2, Message := 'Channel2 on before the error');

// act
group_3(Run := TRUE);
terminal_3(SafeOut1 := TRUE, SafeOut2 := TRUE, InjectComError := TRUE, StartupTime := T#0S);

// assert
AssertEquals_BOOL(Expected := TRUE, Actual := terminal_3.ComError, Message := 'com error');
AssertEquals_BOOL(Expected := FALSE, Actual := terminal_3.Channel1, Message := 'Channel1 fail-safe on com error');
AssertEquals_BOOL(Expected := FALSE, Actual := terminal_3.Channel2, Message := 'Channel2 fail-safe on com error');
TEST_FINISHED_NAMED(__POUNAME());
END_METHOD

METHOD PRIVATE Test_GroupNotRunningForcesChannelsFalse
TcUnit.TEST(__POUNAME());
// arrange: connection in Data with the group running
FOR i_5 := 1 TO 10 DO
    group_5(Run := TRUE, ModuleFault := FALSE);
    terminal_5(StartupTime := T#0S, SafeOut1 := TRUE, SafeOut2 := TRUE);
END_FOR
AssertEquals_BOOL(Expected := TRUE, Actual := terminal_5.Channel1, Message := 'channel on while the group runs');
// act: group STOP (the connection stays in Data)
group_5(Run := FALSE, ModuleFault := FALSE);
terminal_5(StartupTime := T#0S, SafeOut1 := TRUE, SafeOut2 := TRUE);
// assert
AssertEquals_BOOL(Expected := TRUE, Actual := terminal_5.InDataState, Message := 'still in Data');
AssertEquals_BOOL(Expected := FALSE, Actual := terminal_5.Channel1, Message := 'outputs off with the group in STOP');
// act: group ERROR
group_5(Run := TRUE, ModuleFault := TRUE);
terminal_5(StartupTime := T#0S, SafeOut1 := TRUE, SafeOut2 := TRUE);
group_5(Run := TRUE, ModuleFault := TRUE);
terminal_5(StartupTime := T#0S, SafeOut1 := TRUE, SafeOut2 := TRUE);
AssertEquals_BYTE(Expected := TO_BYTE(E_SafeGroupState.Error), Actual := group_5.State, Message := 'group in ERROR');
AssertEquals_BOOL(Expected := FALSE, Actual := terminal_5.Channel2, Message := 'outputs off with the group in ERROR');
TEST_FINISHED_NAMED(__POUNAME());
END_METHOD

METHOD PRIVATE Test_RegistersAsConnection
TcUnit.TEST(__POUNAME());

// act
group_4(Run := TRUE);
terminal_4(StartupTime := T#0S);

// assert
AssertEquals_UINT(Expected := 1, Actual := group_4.ConnectionCount, Message := 'one connection registered');
AssertEquals_UINT(Expected := 0, Actual := group_4.FunctionBlockCount, Message := 'no function blocks');
TEST_FINISHED_NAMED(__POUNAME());
END_METHOD

END_FUNCTION_BLOCK

// Tests/T_SafeConnShutdown_Tests
FUNCTION_BLOCK T_SafeConnShutdown_Tests EXTENDS TcUnit.FB_TestSuite
VAR
    // Test_DeactivateShutsDownConnection
    group_1 : T_SafeGroup;
    conn_1 : T_SafeConnection(group := group_1);
    fb_1 : T_SafeConnShutdown(group := group_1, connection := conn_1);
    i_1 : INT;
END_VAR

Test_DeactivateShutsDownConnection();

METHOD PRIVATE Test_DeactivateShutsDownConnection
TcUnit.TEST(__POUNAME());

// arrange: connection up
FOR i_1 := 1 TO 5 DO
    group_1(Run := TRUE);
    conn_1(StartupTime := T#0S);
    fb_1(Deactivate1 := FALSE);
END_FOR

AssertEquals_BOOL(Expected := FALSE, Actual := fb_1.Deactivated, Message := 'connection up');
// act
group_1(Run := TRUE);
fb_1(Deactivate1 := TRUE);
conn_1(StartupTime := T#0S);
fb_1(Deactivate1 := TRUE);
// assert
AssertEquals_BOOL(Expected := TRUE, Actual := conn_1.IsShutdown, Message := 'connection shut down');
AssertEquals_BOOL(Expected := TRUE, Actual := fb_1.Deactivated, Message := 'Deactivated output on');

// act: release
FOR i_1 := 1 TO 6 DO
    group_1(Run := TRUE);
    fb_1(Deactivate1 := FALSE);
    conn_1(StartupTime := T#0S);
END_FOR

AssertEquals_BOOL(Expected := TRUE, Actual := conn_1.InDataState, Message := 'connection re-established');
AssertEquals_BOOL(Expected := FALSE, Actual := fb_1.Deactivated, Message := 'Deactivated output off');
TEST_FINISHED_NAMED(__POUNAME());
END_METHOD

END_FUNCTION_BLOCK

// Tests/T_SafeGroup_Tests
FUNCTION_BLOCK T_SafeGroup_Tests EXTENDS TcUnit.FB_TestSuite
VAR
    // Test_StopWhenRunFalse
    group_1 : T_SafeGroup;
    fb_1 : T_SafeAnd(group := group_1);
    // Test_RunsFunctionBlocksWithoutConnections
    group_2 : T_SafeGroup;
    fb_2 : T_SafeAnd(group := group_2);
    // Test_FbErrorStopsGroupAndErrAckRecovers
    group_3 : T_SafeGroup;
    eStop_3 : T_SafeEStop(group := group_3);
    andFb_3 : T_SafeAnd(group := group_3);
    // Test_ConnectionStartupAndComError
    group_4 : T_SafeGroup;
    terminal_4 : T_SafeInputTerminal(group := group_4);
    state_4 : INT := 10;
    waitTimer_4 : TON;
    // Test_RegistersMoreThanSixtyFourBlocks
    group_5 : T_SafeGroup;
    blocks_5 : ARRAY[1..70] OF T_SafeAnd(group := group_5);
    // Test_RefusesTheSixtyFifthConnection
    group_6 : T_SafeGroup;
    terminals_6 : ARRAY[1..65] OF T_SafeInputTerminal(group := group_6);
END_VAR

Test_StopWhenRunFalse();
Test_RunsFunctionBlocksWithoutConnections();
Test_FbErrorStopsGroupAndErrAckRecovers();
Test_ConnectionStartupAndComError();
Test_RegistersMoreThanSixtyFourBlocks();
Test_RefusesTheSixtyFifthConnection();

METHOD PRIVATE Test_ConnectionStartupAndComError
TcUnit.TEST(__POUNAME());
waitTimer_4();

CASE state_4 OF
    10:
        // arrange: terminal_4 starting up
        group_4(Run := TRUE, ErrAck := FALSE);
        terminal_4(InjectComError := FALSE, StartupTime := T#150MS);
        group_4(Run := TRUE, ErrAck := FALSE);
        terminal_4(InjectComError := FALSE, StartupTime := T#150MS);
        // assert
        AssertEquals_BYTE(
            Expected := TO_BYTE(E_SafeGroupState.Start),
            Actual := group_4.State,
            Message := 'group START while the connection starts up'
        );

        AssertEquals_BOOL(Expected := TRUE, Actual := group_4.ComStartup, Message := 'ComStartup');
        state_4 := 20;
        waitTimer_4(IN := TRUE, PT := T#400MS);
    20:
        group_4(Run := TRUE, ErrAck := FALSE);
        terminal_4(InjectComError := FALSE, StartupTime := T#150MS);

        IF NOT waitTimer_4.Q THEN
            RETURN;
        END_IF

        waitTimer_4(IN := FALSE);
        AssertEquals_BYTE(Expected := TO_BYTE(E_SafeGroupState.Run), Actual := group_4.State, Message := 'group RUN once the connection is in Data');
        // act: communication error
        group_4(Run := TRUE, ErrAck := FALSE);
        terminal_4(InjectComError := TRUE, StartupTime := T#150MS);
        group_4(Run := TRUE, ErrAck := FALSE);
        terminal_4(InjectComError := FALSE, StartupTime := T#150MS);
        AssertEquals_BOOL(Expected := TRUE, Actual := group_4.ComErr, Message := 'ComErr');
        AssertEquals_BYTE(Expected := TO_BYTE(E_SafeGroupState.Error), Actual := group_4.State, Message := 'group ERROR');
        group_4(Run := TRUE, ErrAck := TRUE);
        terminal_4(InjectComError := FALSE, StartupTime := T#150MS);
        group_4(Run := TRUE, ErrAck := TRUE);
        terminal_4(InjectComError := FALSE, StartupTime := T#150MS);
        AssertEquals_BYTE(Expected := TO_BYTE(E_SafeGroupState.Reset), Actual := group_4.State, Message := 'group RESET');
        group_4(Run := TRUE, ErrAck := FALSE);
        terminal_4(InjectComError := FALSE, StartupTime := T#150MS);
        AssertEquals_BYTE(Expected := TO_BYTE(E_SafeGroupState.Start), Actual := group_4.State, Message := 'group START again after ack');
        state_4 := 30;
        waitTimer_4(IN := TRUE, PT := T#400MS);
    30:
        group_4(Run := TRUE, ErrAck := FALSE);
        terminal_4(InjectComError := FALSE, StartupTime := T#150MS);

        IF NOT waitTimer_4.Q THEN
            RETURN;
        END_IF

        waitTimer_4(IN := FALSE);
        AssertEquals_BYTE(Expected := TO_BYTE(E_SafeGroupState.Run), Actual := group_4.State, Message := 'group RUN after reconnection');
        TEST_FINISHED_NAMED(__POUNAME());
        state_4 := 10;
END_CASE
END_METHOD

METHOD PRIVATE Test_FbErrorStopsGroupAndErrAckRecovers
TcUnit.TEST(__POUNAME());
// arrange: an AND that runs and an ESTOP that will raise an EDM error
group_3(Run := TRUE, ErrAck := FALSE);
eStop_3(Restart := FALSE, EDM1 := FALSE, EStopIn1 := TRUE);
andFb_3(AndIn1 := TRUE, AndIn2 := TRUE);
group_3(Run := TRUE, ErrAck := FALSE);
eStop_3(Restart := FALSE, EDM1 := FALSE, EStopIn1 := TRUE);
andFb_3(AndIn1 := TRUE, AndIn2 := TRUE);
AssertEquals_BOOL(Expected := TRUE, Actual := andFb_3.AndOut, Message := 'AND running before the error');
// act: restart with missing feedback -> FB error
group_3(Run := TRUE, ErrAck := FALSE);
eStop_3(Restart := TRUE, EDM1 := FALSE, EStopIn1 := TRUE);
andFb_3(AndIn1 := TRUE, AndIn2 := TRUE);
group_3(Run := TRUE, ErrAck := FALSE);
eStop_3(Restart := FALSE, EDM1 := FALSE, EStopIn1 := TRUE);
andFb_3(AndIn1 := TRUE, AndIn2 := TRUE);
// assert
AssertEquals_BOOL(Expected := TRUE, Actual := group_3.FbErr, Message := 'FbErr');
AssertEquals_BYTE(Expected := TO_BYTE(E_SafeGroupState.Error), Actual := group_3.State, Message := 'group ERROR');
AssertEquals_BYTE(Expected := TO_BYTE(E_SafeGroupDiag.FbError), Actual := group_3.Diag, Message := 'group diag FBERROR');
AssertEquals_BOOL(Expected := FALSE, Actual := andFb_3.AndOut, Message := 'other FB outputs forced safe');
AssertEquals_BYTE(Expected := TO_BYTE(E_SafeFbState.Stop), Actual := andFb_3.State, Message := 'other FB STOP');
// act: ErrAck 0 -> 1 -> 0
group_3(Run := TRUE, ErrAck := TRUE);
eStop_3(Restart := FALSE, EDM1 := FALSE, EStopIn1 := TRUE);
andFb_3(AndIn1 := TRUE, AndIn2 := TRUE);
group_3(Run := TRUE, ErrAck := TRUE);
eStop_3(Restart := FALSE, EDM1 := FALSE, EStopIn1 := TRUE);
andFb_3(AndIn1 := TRUE, AndIn2 := TRUE);
AssertEquals_BYTE(Expected := TO_BYTE(E_SafeGroupState.Reset), Actual := group_3.State, Message := 'group RESET while ErrAck 1');
group_3(Run := TRUE, ErrAck := FALSE);
eStop_3(Restart := FALSE, EDM1 := FALSE, EStopIn1 := TRUE);
andFb_3(AndIn1 := TRUE, AndIn2 := TRUE);
group_3(Run := TRUE, ErrAck := FALSE);
eStop_3(Restart := FALSE, EDM1 := FALSE, EStopIn1 := TRUE);
andFb_3(AndIn1 := TRUE, AndIn2 := TRUE);
AssertEquals_BYTE(Expected := TO_BYTE(E_SafeGroupState.Run), Actual := group_3.State, Message := 'group RUN after ErrAck');
AssertEquals_BOOL(Expected := TRUE, Actual := andFb_3.AndOut, Message := 'AND running again');
AssertEquals_BYTE(Expected := TO_BYTE(E_SafeFbState.Safe), Actual := eStop_3.State, Message := 'ESTOP back in SAFE awaiting restart');
TEST_FINISHED_NAMED(__POUNAME());
END_METHOD

METHOD PRIVATE Test_RefusesTheSixtyFifthConnection
TcUnit.TEST(__POUNAME());
// arrange: 65 terminals tried to join group_6 at initialisation
// assert
AssertEquals_UINT(Expected := 64, Actual := group_6.ConnectionCount, Message := 'the cap holds');
AssertEquals_BOOL(Expected := TRUE, Actual := group_6.RegistrationRefused, Message := 'the refusal is visible');
TEST_FINISHED_NAMED(__POUNAME());
END_METHOD

METHOD PRIVATE Test_RegistersMoreThanSixtyFourBlocks
TcUnit.TEST(__POUNAME());
// arrange: 70 blocks joined group_5 at initialisation
// assert
AssertEquals_UINT(Expected := 70, Actual := group_5.FunctionBlockCount, Message := 'every block registered');
AssertEquals_BOOL(Expected := FALSE, Actual := group_5.RegistrationRefused, Message := 'none refused');
TEST_FINISHED_NAMED(__POUNAME());
END_METHOD

METHOD PRIVATE Test_RunsFunctionBlocksWithoutConnections
TcUnit.TEST(__POUNAME());
// act
group_2(Run := TRUE);
fb_2(AndIn1 := TRUE, AndIn2 := TRUE);
group_2(Run := TRUE);
fb_2(AndIn1 := TRUE, AndIn2 := TRUE);
// assert
AssertEquals_BYTE(Expected := TO_BYTE(E_SafeGroupState.Run), Actual := group_2.State, Message := 'group RUN');
AssertEquals_BOOL(Expected := TRUE, Actual := fb_2.AndOut, Message := 'FB executed');
AssertEquals_BOOL(Expected := TRUE, Actual := group_2.FbRun, Message := 'all FBs running');
TEST_FINISHED_NAMED(__POUNAME());
END_METHOD

METHOD PRIVATE Test_StopWhenRunFalse
TcUnit.TEST(__POUNAME());
// act
group_1(Run := FALSE);
fb_1(AndIn1 := TRUE, AndIn2 := TRUE);
// assert
AssertEquals_BYTE(Expected := TO_BYTE(E_SafeGroupState.Stop), Actual := group_1.State, Message := 'group STOP');
AssertEquals_BYTE(Expected := TO_BYTE(E_SafeFbState.Stop), Actual := fb_1.State, Message := 'FB STOP');
AssertEquals_BOOL(Expected := FALSE, Actual := group_1.InRun, Message := 'InRun off');
TEST_FINISHED_NAMED(__POUNAME());
END_METHOD

END_FUNCTION_BLOCK

// Tests/T_SafeAnd_Tests_CFC
    // CFC twin of T_SafeAnd_Tests: the same tests drawn as CFC diagrams, the way a TwinSAFE project is authored.
    FUNCTION_BLOCK T_SafeAnd_Tests_CFC EXTENDS T_SafeCfcTestSuite
    VAR
    // Test_AllConnectedInputsTrueGivesRun
    group_1 : T_SafeGroup;
    fb_1 : T_SafeAnd(group := group_1);
    // Test_OneInputFalseGivesSafe
    group_2 : T_SafeGroup;
    fb_2 : T_SafeAnd(group := group_2);
    // Test_UnconnectedInputsIgnoredAndMakeContactNegated
    group_3 : T_SafeGroup;
    fb_3 : T_SafeAnd(group := group_3) := (Parameters := (In2MakeContact := TRUE));
    // Test_StoppedGivesNoOutput
    group_4 : T_SafeGroup;
    fb_4 : T_SafeAnd(group := group_4);
END_VAR

Test_AllConnectedInputsTrueGivesRun();
Test_OneInputFalseGivesSafe();
Test_UnconnectedInputsIgnoredAndMakeContactNegated();
Test_StoppedGivesNoOutput();

METHOD PRIVATE Test_AllConnectedInputsTrueGivesRun
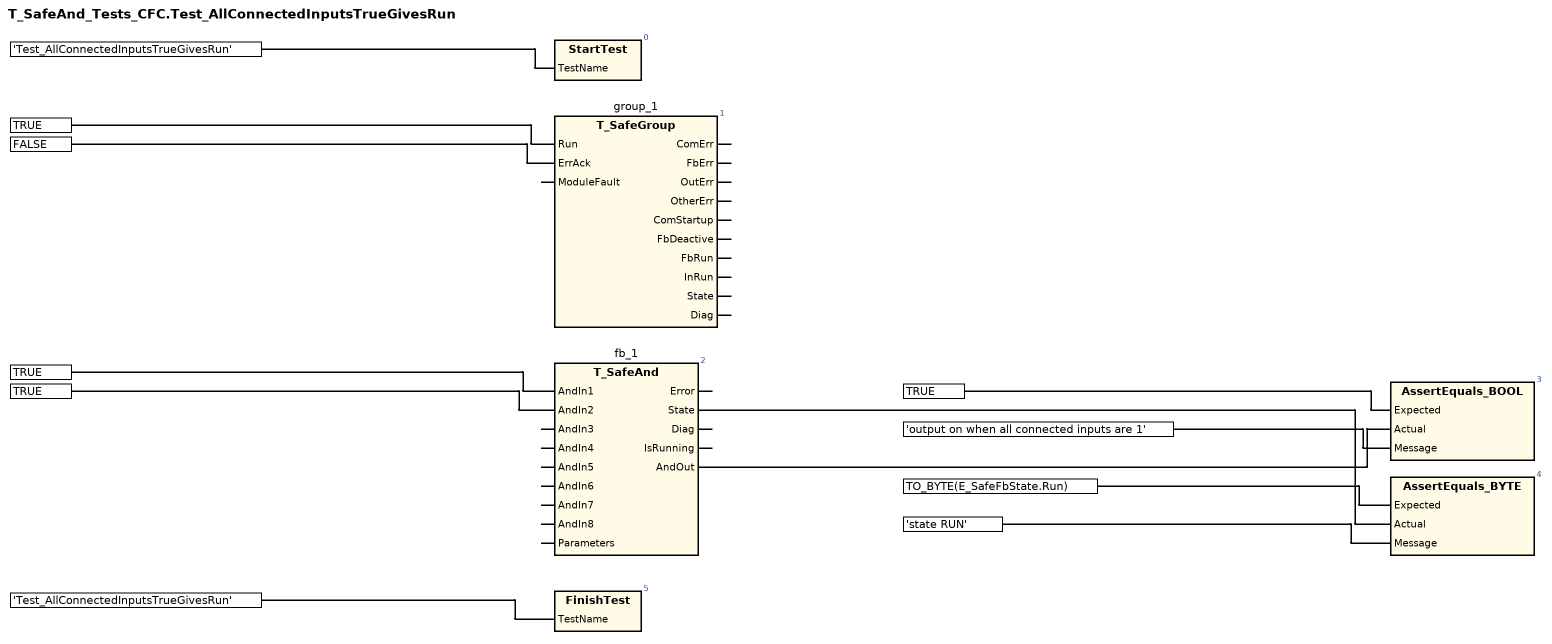
StartTest(TestName := 'Test_AllConnectedInputsTrueGivesRun');
group_1(Run := TRUE, ErrAck := FALSE); // T_SafeGroup
fb_1(AndIn1 := TRUE, AndIn2 := TRUE); // T_SafeAnd
AssertEquals_BOOL(Expected := TRUE, Actual := fb_1.AndOut, Message := 'output on when all connected inputs are 1');
AssertEquals_BYTE(Expected := TO_BYTE(E_SafeFbState.Run), Actual := fb_1.State, Message := 'state RUN');
FinishTest(TestName := 'Test_AllConnectedInputsTrueGivesRun');
END_METHOD

METHOD PRIVATE Test_OneInputFalseGivesSafe
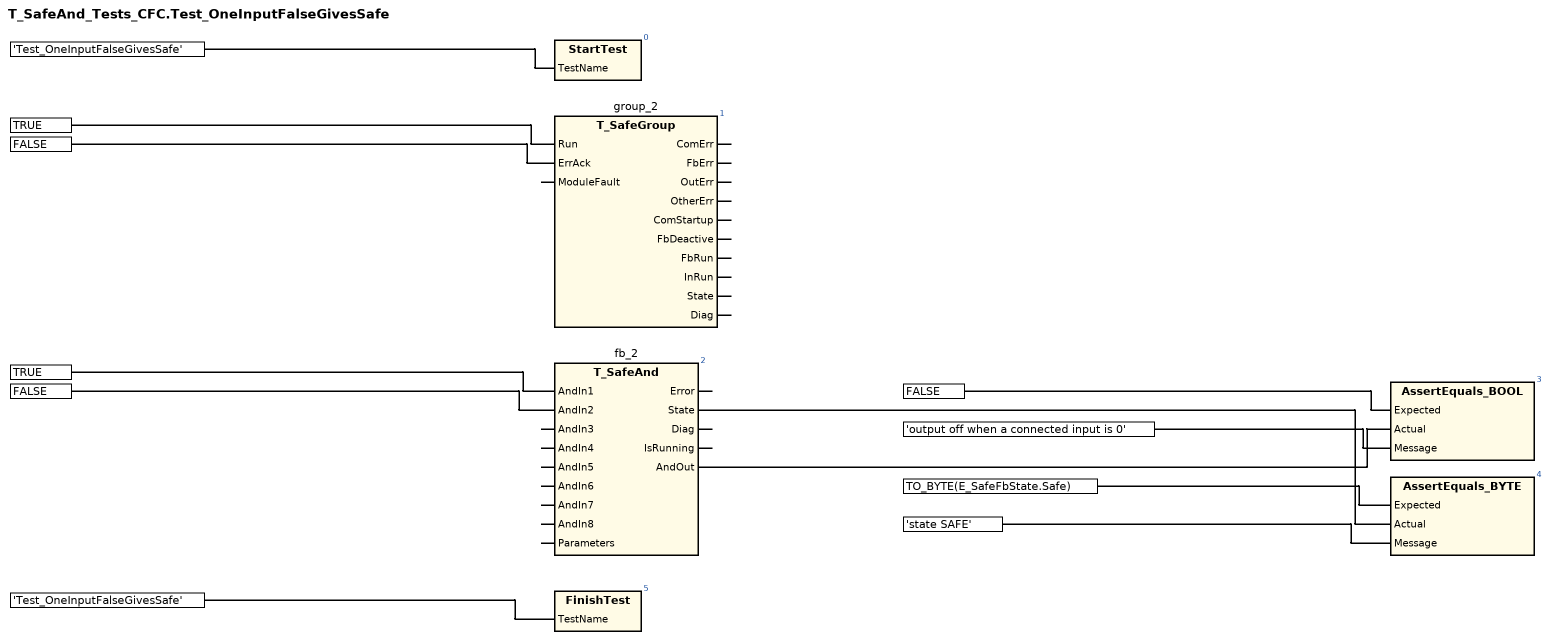
StartTest(TestName := 'Test_OneInputFalseGivesSafe');
group_2(Run := TRUE, ErrAck := FALSE); // T_SafeGroup
fb_2(AndIn1 := TRUE, AndIn2 := FALSE); // T_SafeAnd
AssertEquals_BOOL(Expected := FALSE, Actual := fb_2.AndOut, Message := 'output off when a connected input is 0');
AssertEquals_BYTE(Expected := TO_BYTE(E_SafeFbState.Safe), Actual := fb_2.State, Message := 'state SAFE');
FinishTest(TestName := 'Test_OneInputFalseGivesSafe');
END_METHOD

METHOD PRIVATE Test_StoppedGivesNoOutput
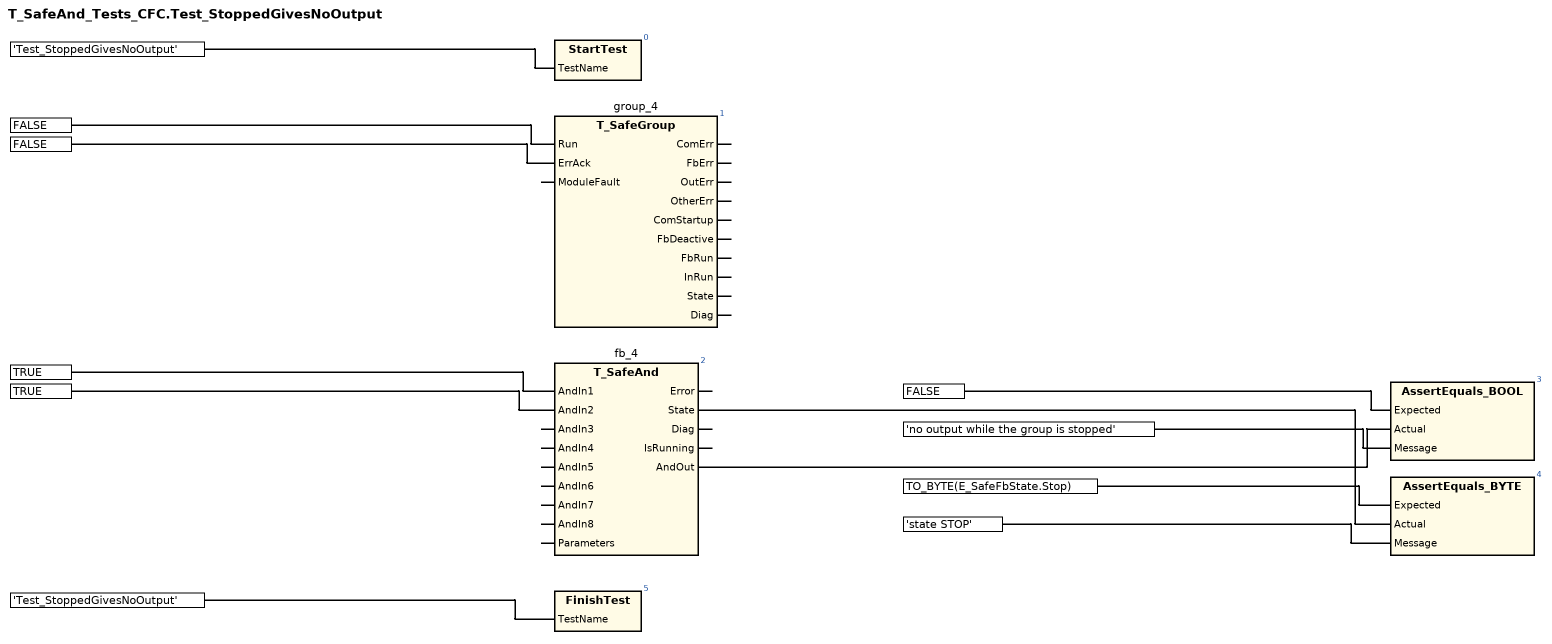
StartTest(TestName := 'Test_StoppedGivesNoOutput');
group_4(Run := FALSE, ErrAck := FALSE); // T_SafeGroup
fb_4(AndIn1 := TRUE, AndIn2 := TRUE); // T_SafeAnd
AssertEquals_BOOL(Expected := FALSE, Actual := fb_4.AndOut, Message := 'no output while the group is stopped');
AssertEquals_BYTE(Expected := TO_BYTE(E_SafeFbState.Stop), Actual := fb_4.State, Message := 'state STOP');
FinishTest(TestName := 'Test_StoppedGivesNoOutput');
END_METHOD

METHOD PRIVATE Test_UnconnectedInputsIgnoredAndMakeContactNegated
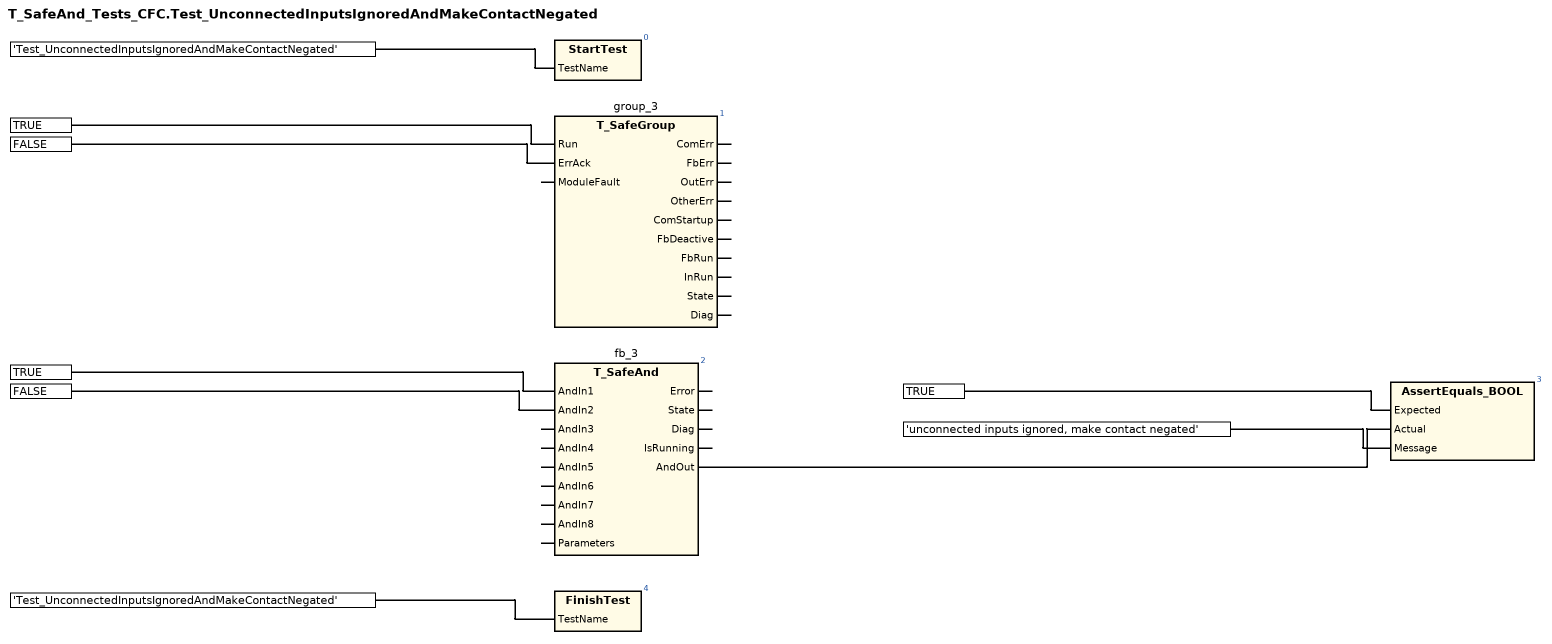
StartTest(TestName := 'Test_UnconnectedInputsIgnoredAndMakeContactNegated');
group_3(Run := TRUE, ErrAck := FALSE); // T_SafeGroup
fb_3(AndIn1 := TRUE, AndIn2 := FALSE); // T_SafeAnd
AssertEquals_BOOL(Expected := TRUE, Actual := fb_3.AndOut, Message := 'unconnected inputs ignored, make contact negated');
FinishTest(TestName := 'Test_UnconnectedInputsIgnoredAndMakeContactNegated');
END_METHOD

END_FUNCTION_BLOCK

// Tests/T_SafeInputPair_Tests_CFC
    // CFC twin of T_SafeInputPair_Tests: the same tests drawn as CFC diagrams, the way a TwinSAFE project is authored.
    FUNCTION_BLOCK T_SafeInputPair_Tests_CFC EXTENDS T_SafeCfcTestSuite
    VAR
    // Test_InactivePairNeverRequestsSafeState
    pair_1 : T_SafeInputPair;
    // Test_BreakContactRequestsSafeStateOnZero
    pair_2 : T_SafeInputPair;
    // Test_MakeContactRequestsSafeStateOnOne
    pair_3 : T_SafeInputPair;
    // Test_TwoChannelRequestsSafeStateIfEitherChannelLow
    pair_4 : T_SafeInputPair;
    // Test_DiscrepancyErrorAfterTimeoutAndResetAfterSafeInputs
    pair_5 : T_SafeInputPair;
    t1_5 : TON;
    t2_5 : TON;
    trig1_5 : R_TRIG;
    trig2_5 : R_TRIG;
END_VAR

Test_InactivePairNeverRequestsSafeState();
Test_BreakContactRequestsSafeStateOnZero();
Test_MakeContactRequestsSafeStateOnOne();
Test_TwoChannelRequestsSafeStateIfEitherChannelLow();
Test_DiscrepancyErrorAfterTimeoutAndResetAfterSafeInputs();

METHOD PRIVATE Test_BreakContactRequestsSafeStateOnZero
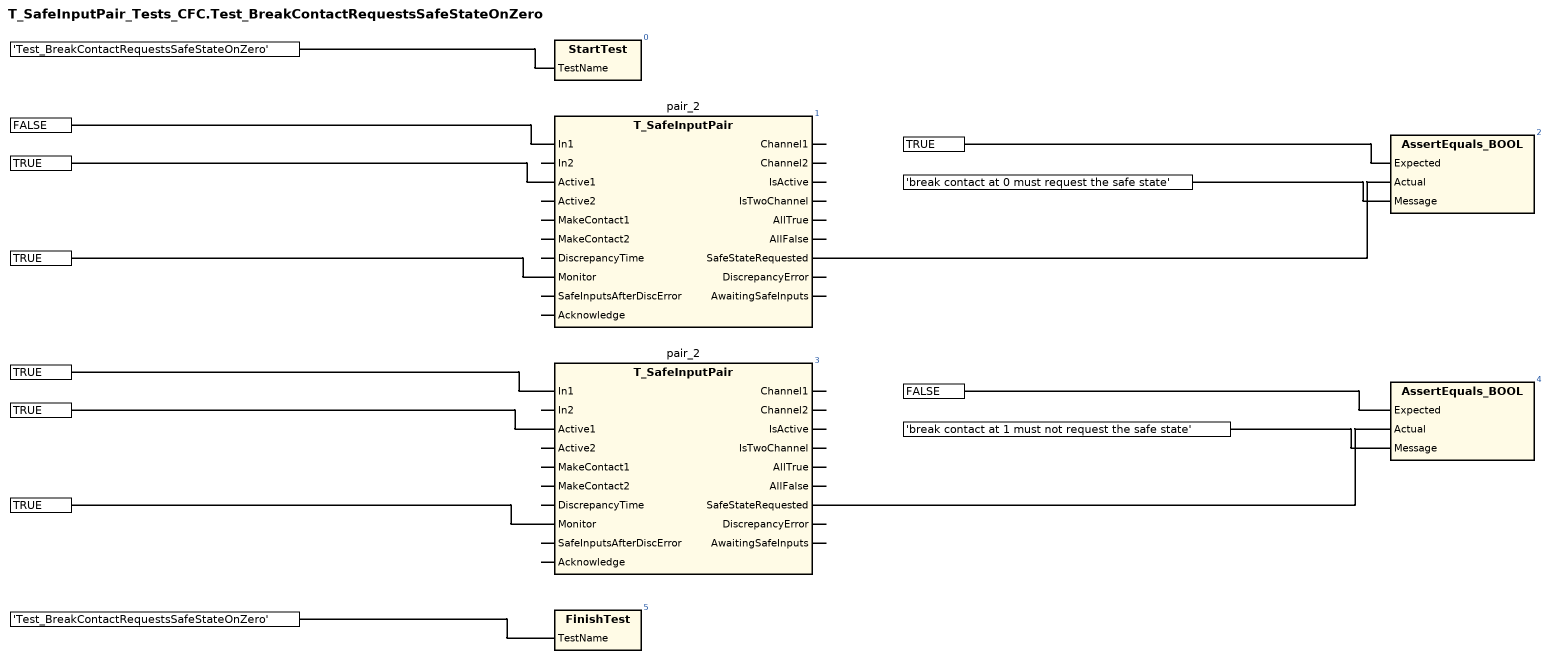
StartTest(TestName := 'Test_BreakContactRequestsSafeStateOnZero');
pair_2(In1 := FALSE, Active1 := TRUE, Monitor := TRUE); // T_SafeInputPair
AssertEquals_BOOL(Expected := TRUE, Actual := pair_2.SafeStateRequested, Message := 'break contact at 0 must request the safe state');
pair_2(In1 := TRUE, Active1 := TRUE, Monitor := TRUE); // T_SafeInputPair
AssertEquals_BOOL(Expected := FALSE, Actual := pair_2.SafeStateRequested, Message := 'break contact at 1 must not request the safe state');
FinishTest(TestName := 'Test_BreakContactRequestsSafeStateOnZero');
END_METHOD

METHOD PRIVATE Test_DiscrepancyErrorAfterTimeoutAndResetAfterSafeInputs
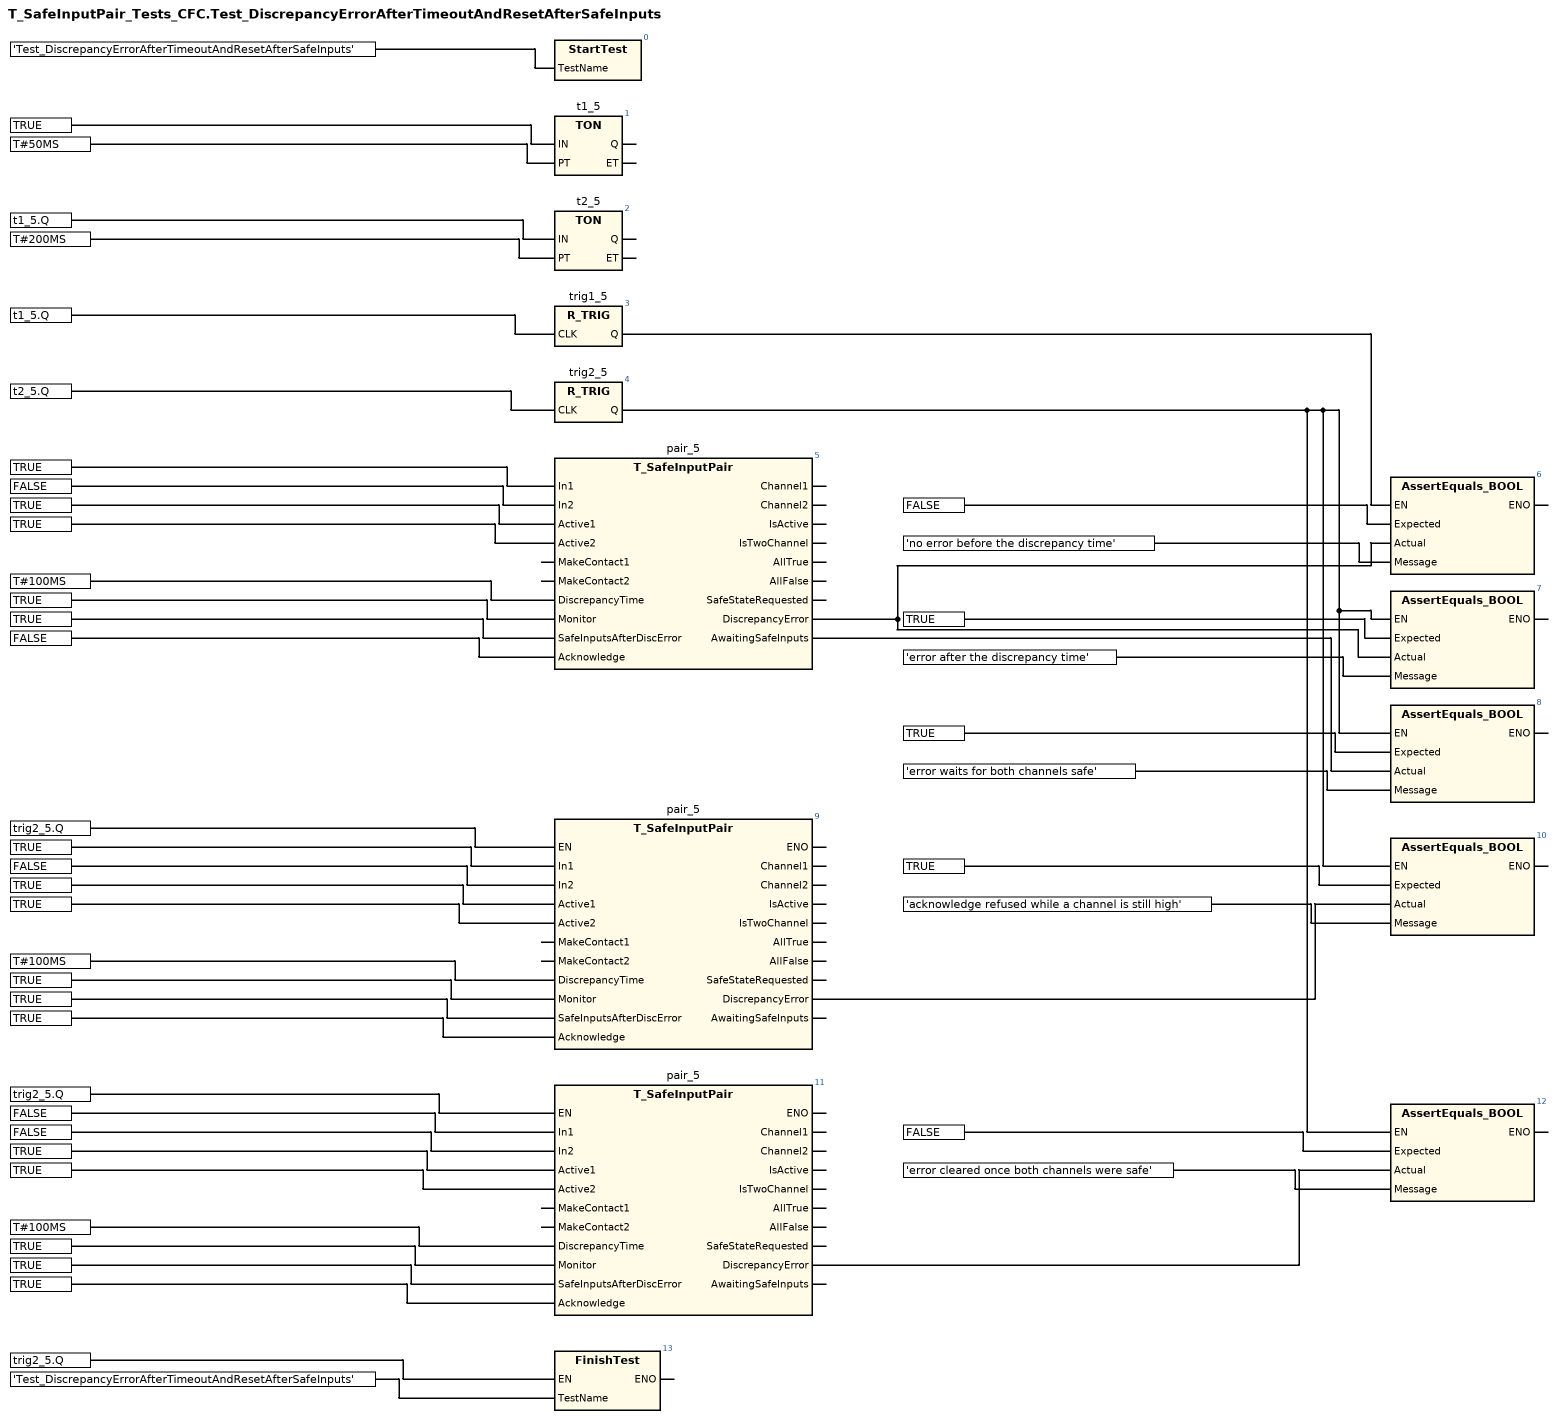
StartTest(TestName := 'Test_DiscrepancyErrorAfterTimeoutAndResetAfterSafeInputs');
t1_5(IN := TRUE, PT := T#50MS); // TON
t2_5(IN := t1_5.Q, PT := T#200MS); // TON
trig1_5(CLK := t1_5.Q); // R_TRIG
trig2_5(CLK := t2_5.Q); // R_TRIG
pair_5(
    In1 := TRUE,
    In2 := FALSE,
    Active1 := TRUE,
    Active2 := TRUE,
    DiscrepancyTime := T#100MS,
    Monitor := TRUE,
    SafeInputsAfterDiscError := TRUE,
    Acknowledge := FALSE); // T_SafeInputPair
IF trig1_5.Q THEN AssertEquals_BOOL(Expected := FALSE, Actual := pair_5.DiscrepancyError, Message := 'no error before the discrepancy time'); END_IF
IF trig2_5.Q THEN AssertEquals_BOOL(Expected := TRUE, Actual := pair_5.DiscrepancyError, Message := 'error after the discrepancy time'); END_IF
IF trig2_5.Q THEN AssertEquals_BOOL(Expected := TRUE, Actual := pair_5.AwaitingSafeInputs, Message := 'error waits for both channels safe'); END_IF
IF trig2_5.Q THEN
    pair_5(
        In1 := TRUE,
        In2 := FALSE,
        Active1 := TRUE,
        Active2 := TRUE,
        DiscrepancyTime := T#100MS,
        Monitor := TRUE,
        SafeInputsAfterDiscError := TRUE,
        Acknowledge := TRUE); // T_SafeInputPair
END_IF
IF trig2_5.Q THEN AssertEquals_BOOL(Expected := TRUE, Actual := pair_5.DiscrepancyError, Message := 'acknowledge refused while a channel is still high'); END_IF
IF trig2_5.Q THEN
    pair_5(
        In1 := FALSE,
        In2 := FALSE,
        Active1 := TRUE,
        Active2 := TRUE,
        DiscrepancyTime := T#100MS,
        Monitor := TRUE,
        SafeInputsAfterDiscError := TRUE,
        Acknowledge := TRUE); // T_SafeInputPair
END_IF
IF trig2_5.Q THEN AssertEquals_BOOL(Expected := FALSE, Actual := pair_5.DiscrepancyError, Message := 'error cleared once both channels were safe'); END_IF
IF trig2_5.Q THEN FinishTest(TestName := 'Test_DiscrepancyErrorAfterTimeoutAndResetAfterSafeInputs'); END_IF
END_METHOD

METHOD PRIVATE Test_InactivePairNeverRequestsSafeState
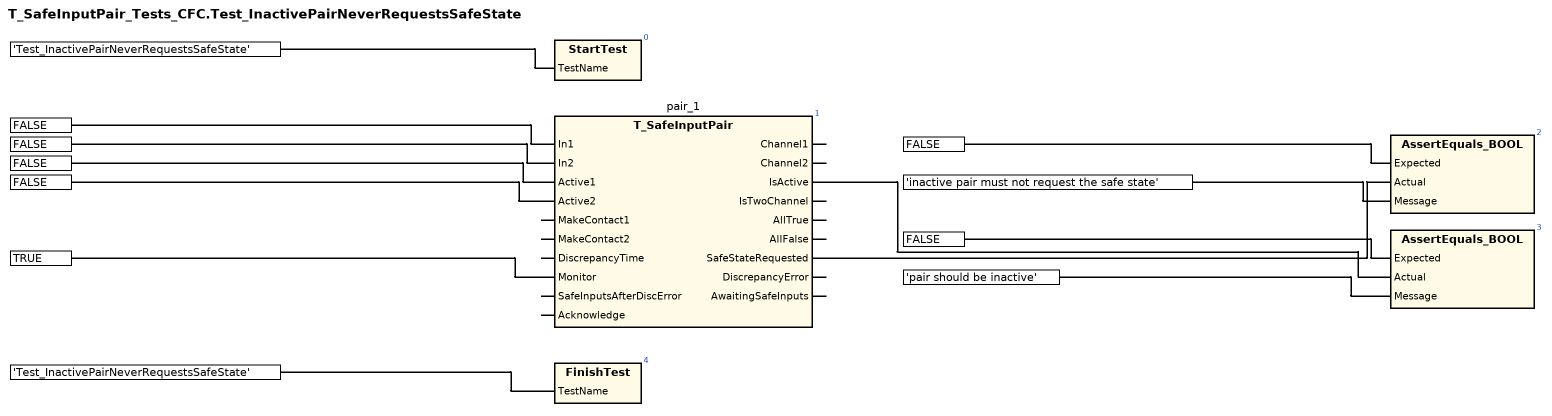
StartTest(TestName := 'Test_InactivePairNeverRequestsSafeState');
pair_1(In1 := FALSE, In2 := FALSE, Active1 := FALSE, Active2 := FALSE, Monitor := TRUE); // T_SafeInputPair
AssertEquals_BOOL(Expected := FALSE, Actual := pair_1.SafeStateRequested, Message := 'inactive pair must not request the safe state');
AssertEquals_BOOL(Expected := FALSE, Actual := pair_1.IsActive, Message := 'pair should be inactive');
FinishTest(TestName := 'Test_InactivePairNeverRequestsSafeState');
END_METHOD

METHOD PRIVATE Test_MakeContactRequestsSafeStateOnOne
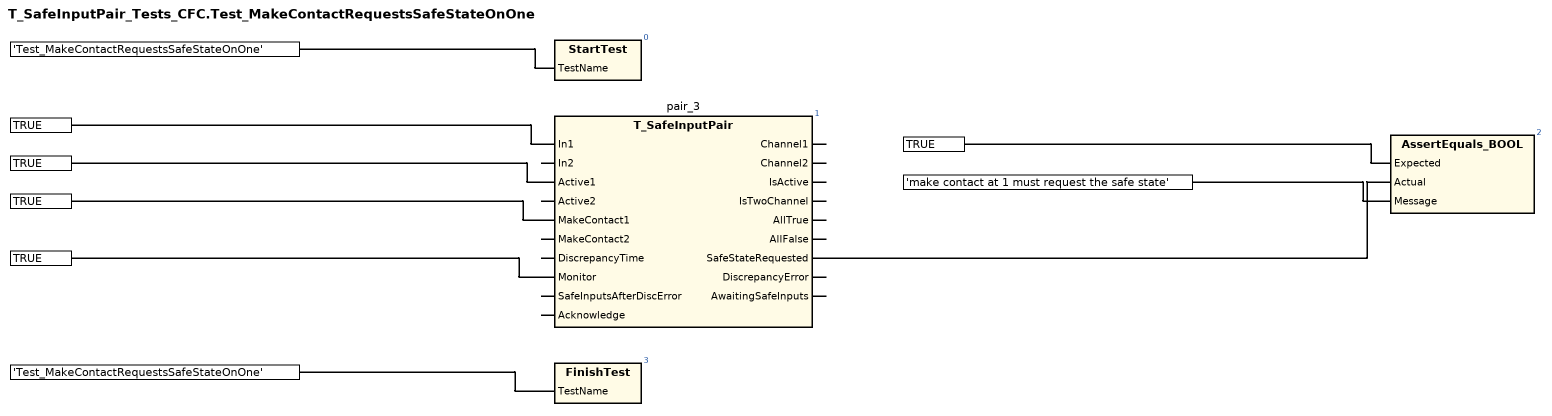
StartTest(TestName := 'Test_MakeContactRequestsSafeStateOnOne');
pair_3(In1 := TRUE, Active1 := TRUE, MakeContact1 := TRUE, Monitor := TRUE); // T_SafeInputPair
AssertEquals_BOOL(Expected := TRUE, Actual := pair_3.SafeStateRequested, Message := 'make contact at 1 must request the safe state');
FinishTest(TestName := 'Test_MakeContactRequestsSafeStateOnOne');
END_METHOD

METHOD PRIVATE Test_TwoChannelRequestsSafeStateIfEitherChannelLow
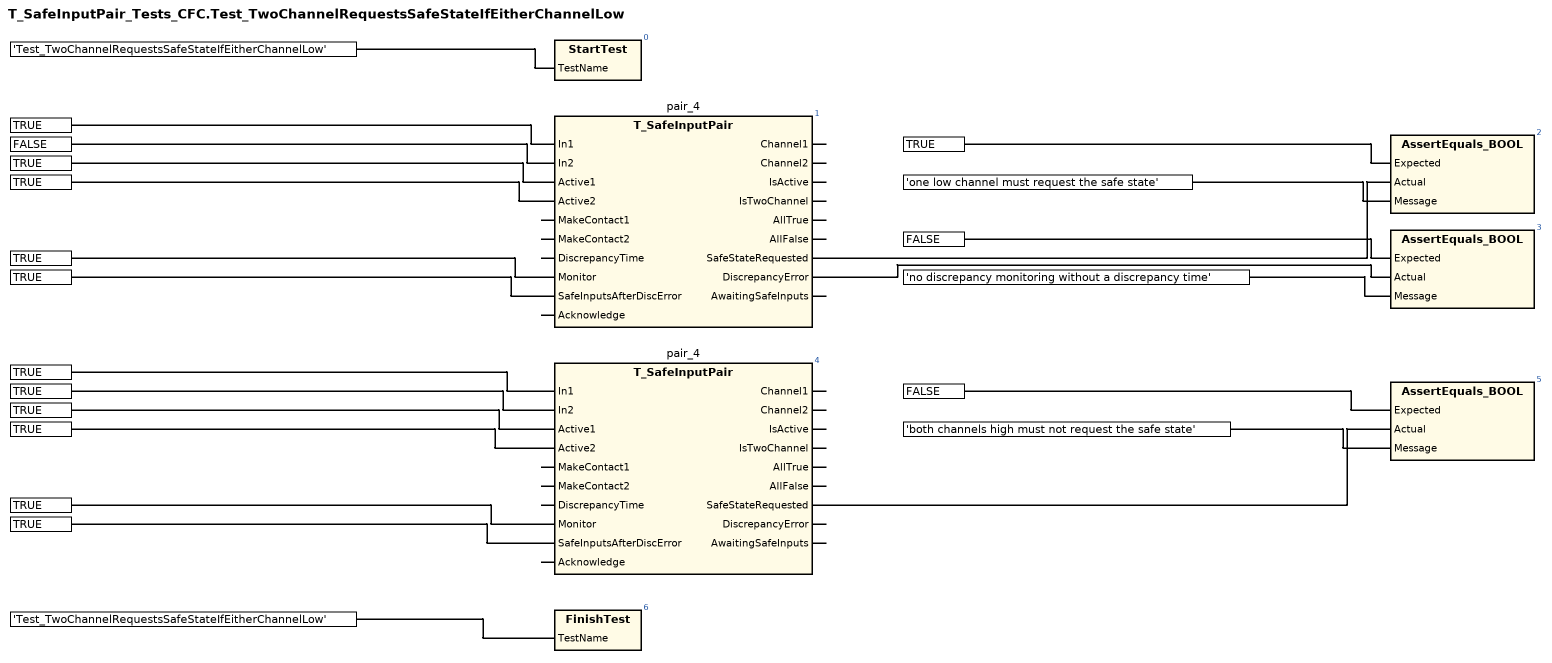
StartTest(TestName := 'Test_TwoChannelRequestsSafeStateIfEitherChannelLow');
pair_4(
    In1 := TRUE,
    In2 := FALSE,
    Active1 := TRUE,
    Active2 := TRUE,
    Monitor := TRUE,
    SafeInputsAfterDiscError := TRUE); // T_SafeInputPair
AssertEquals_BOOL(Expected := TRUE, Actual := pair_4.SafeStateRequested, Message := 'one low channel must request the safe state');
AssertEquals_BOOL(Expected := FALSE, Actual := pair_4.DiscrepancyError, Message := 'no discrepancy monitoring without a discrepancy time');
pair_4(
    In1 := TRUE,
    In2 := TRUE,
    Active1 := TRUE,
    Active2 := TRUE,
    Monitor := TRUE,
    SafeInputsAfterDiscError := TRUE); // T_SafeInputPair
AssertEquals_BOOL(Expected := FALSE, Actual := pair_4.SafeStateRequested, Message := 'both channels high must not request the safe state');
FinishTest(TestName := 'Test_TwoChannelRequestsSafeStateIfEitherChannelLow');
END_METHOD

END_FUNCTION_BLOCK

// Tests/T_SafeOr_Tests_CFC
    // CFC twin of T_SafeOr_Tests: the same tests drawn as CFC diagrams, the way a TwinSAFE project is authored.
    FUNCTION_BLOCK T_SafeOr_Tests_CFC EXTENDS T_SafeCfcTestSuite
    VAR
    // Test_AnyConnectedInputTrueGivesRun
    group_1 : T_SafeGroup;
    fb_1 : T_SafeOr(group := group_1);
    // Test_AllFalseGivesSafe
    group_2 : T_SafeGroup;
    fb_2 : T_SafeOr(group := group_2);
END_VAR

Test_AnyConnectedInputTrueGivesRun();
Test_AllFalseGivesSafe();

METHOD PRIVATE Test_AllFalseGivesSafe
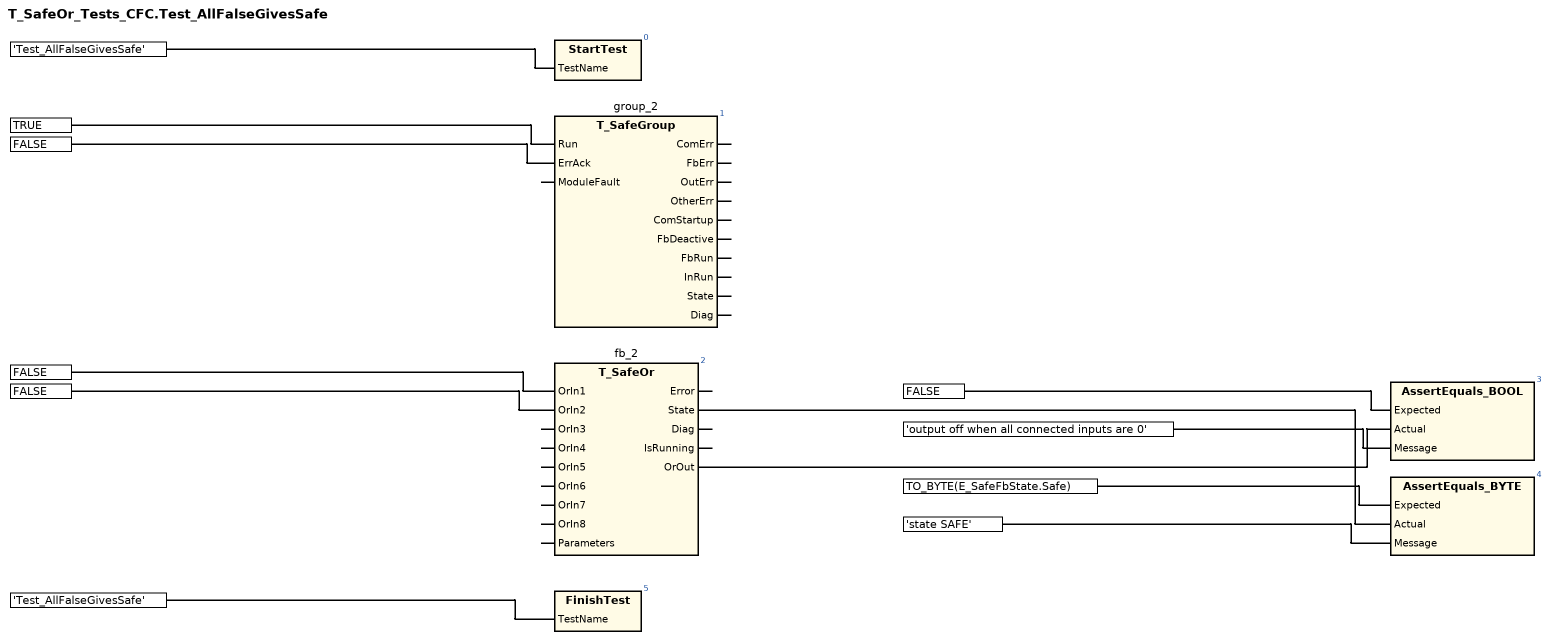
StartTest(TestName := 'Test_AllFalseGivesSafe');
group_2(Run := TRUE, ErrAck := FALSE); // T_SafeGroup
fb_2(OrIn1 := FALSE, OrIn2 := FALSE); // T_SafeOr
AssertEquals_BOOL(Expected := FALSE, Actual := fb_2.OrOut, Message := 'output off when all connected inputs are 0');
AssertEquals_BYTE(Expected := TO_BYTE(E_SafeFbState.Safe), Actual := fb_2.State, Message := 'state SAFE');
FinishTest(TestName := 'Test_AllFalseGivesSafe');
END_METHOD

METHOD PRIVATE Test_AnyConnectedInputTrueGivesRun
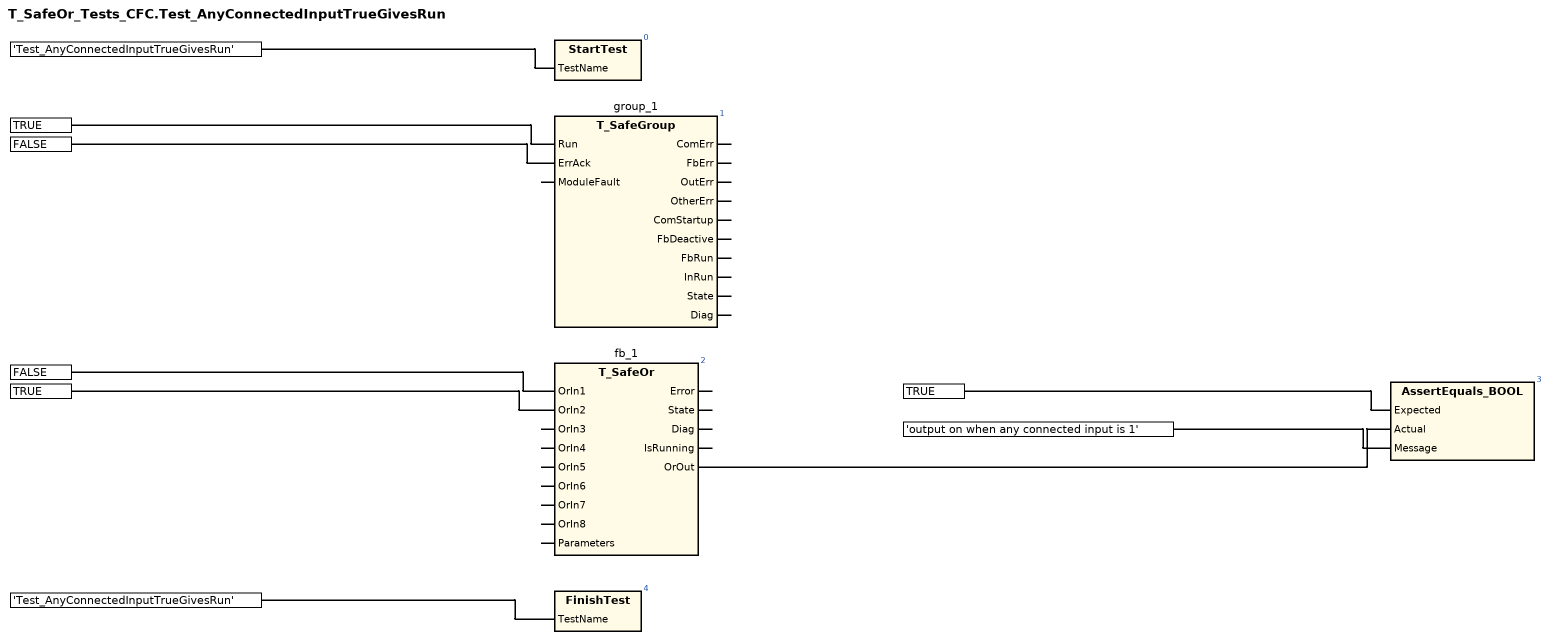
StartTest(TestName := 'Test_AnyConnectedInputTrueGivesRun');
group_1(Run := TRUE, ErrAck := FALSE); // T_SafeGroup
fb_1(OrIn1 := FALSE, OrIn2 := TRUE); // T_SafeOr
AssertEquals_BOOL(Expected := TRUE, Actual := fb_1.OrOut, Message := 'output on when any connected input is 1');
FinishTest(TestName := 'Test_AnyConnectedInputTrueGivesRun');
END_METHOD

END_FUNCTION_BLOCK

// Tests/T_SafeXor_Tests_CFC
    // CFC twin of T_SafeXor_Tests: the same tests drawn as CFC diagrams, the way a TwinSAFE project is authored.
    FUNCTION_BLOCK T_SafeXor_Tests_CFC EXTENDS T_SafeCfcTestSuite
    VAR
    // Test_ConnectedPairsAreExclusiveOr
    group_1 : T_SafeGroup;
    fb_1 : T_SafeXor(group := group_1);
END_VAR

Test_ConnectedPairsAreExclusiveOr();

METHOD PRIVATE Test_ConnectedPairsAreExclusiveOr
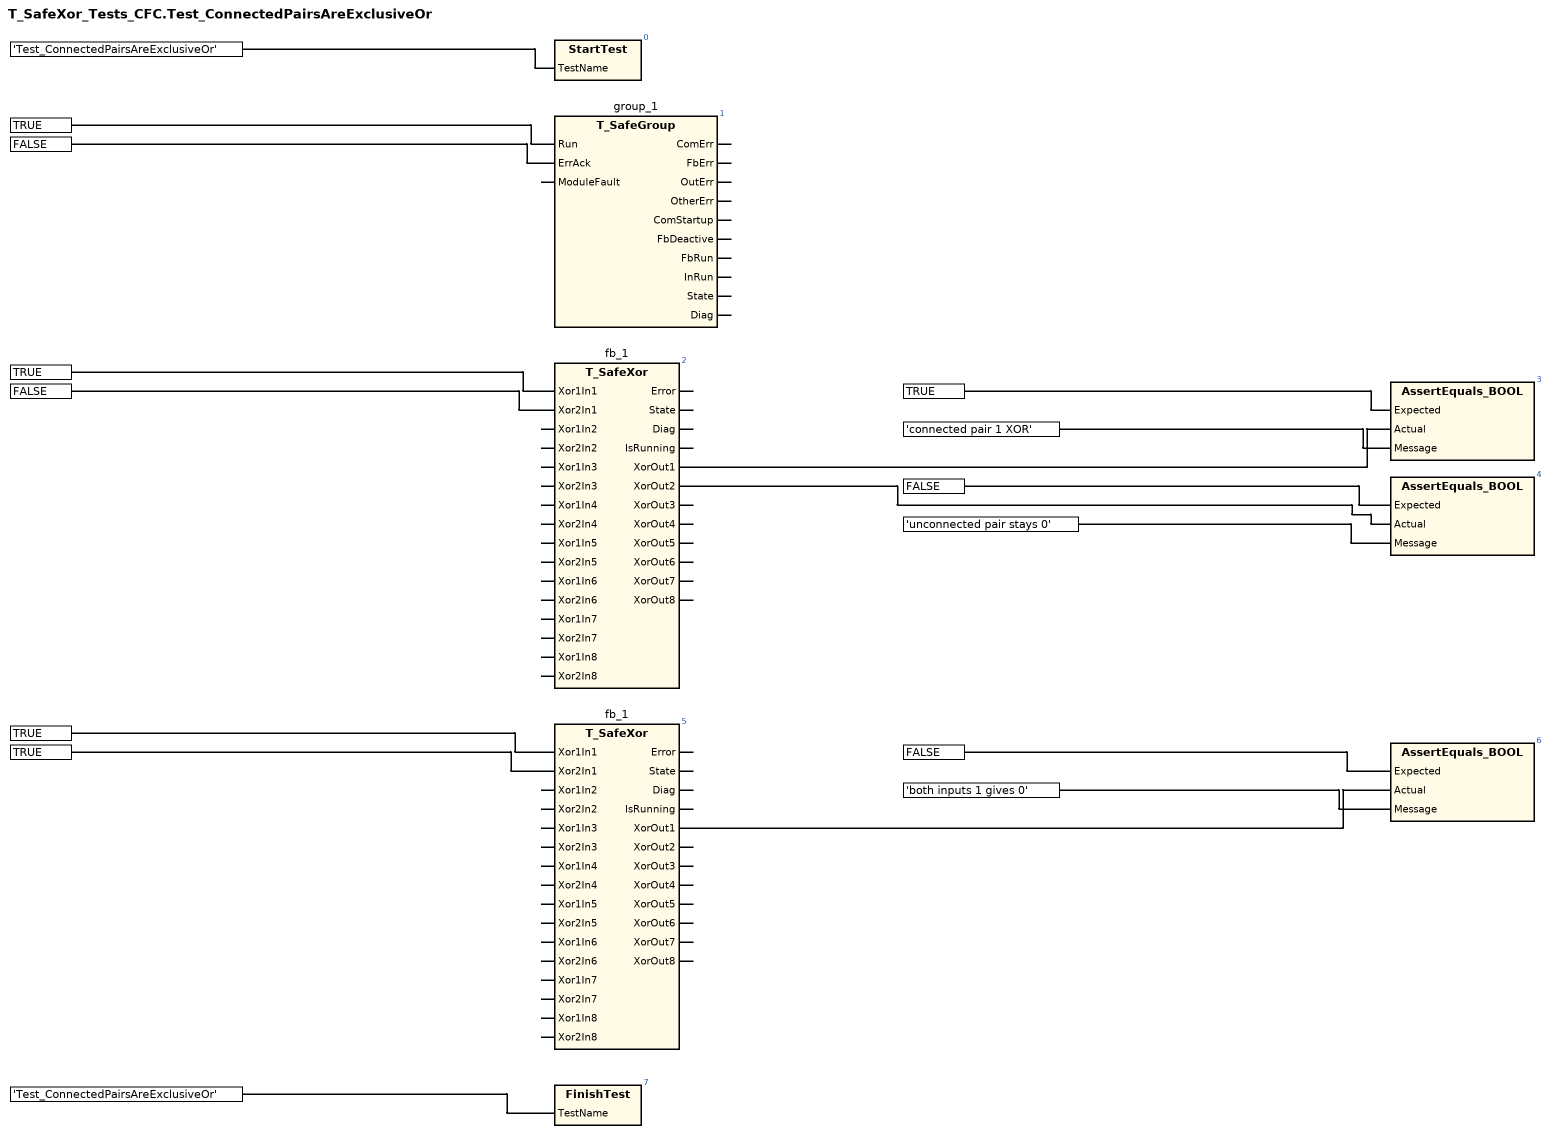
StartTest(TestName := 'Test_ConnectedPairsAreExclusiveOr');
group_1(Run := TRUE, ErrAck := FALSE); // T_SafeGroup
fb_1(Xor1In1 := TRUE, Xor2In1 := FALSE); // T_SafeXor
AssertEquals_BOOL(Expected := TRUE, Actual := fb_1.XorOut1, Message := 'connected pair 1 XOR');
AssertEquals_BOOL(Expected := FALSE, Actual := fb_1.XorOut2, Message := 'unconnected pair stays 0');
fb_1(Xor1In1 := TRUE, Xor2In1 := TRUE); // T_SafeXor
AssertEquals_BOOL(Expected := FALSE, Actual := fb_1.XorOut1, Message := 'both inputs 1 gives 0');
FinishTest(TestName := 'Test_ConnectedPairsAreExclusiveOr');
END_METHOD

END_FUNCTION_BLOCK

// Tests/T_SafeDecouple_Tests_CFC
    // CFC twin of T_SafeDecouple_Tests: the same tests drawn as CFC diagrams, the way a TwinSAFE project is authored.
    FUNCTION_BLOCK T_SafeDecouple_Tests_CFC EXTENDS T_SafeCfcTestSuite
    VAR
    // Test_InputsLoopedToOutputsOnlyWhenRunning
    group_1 : T_SafeGroup;
    fb_1 : T_SafeDecouple(group := group_1);
END_VAR

Test_InputsLoopedToOutputsOnlyWhenRunning();

METHOD PRIVATE Test_InputsLoopedToOutputsOnlyWhenRunning
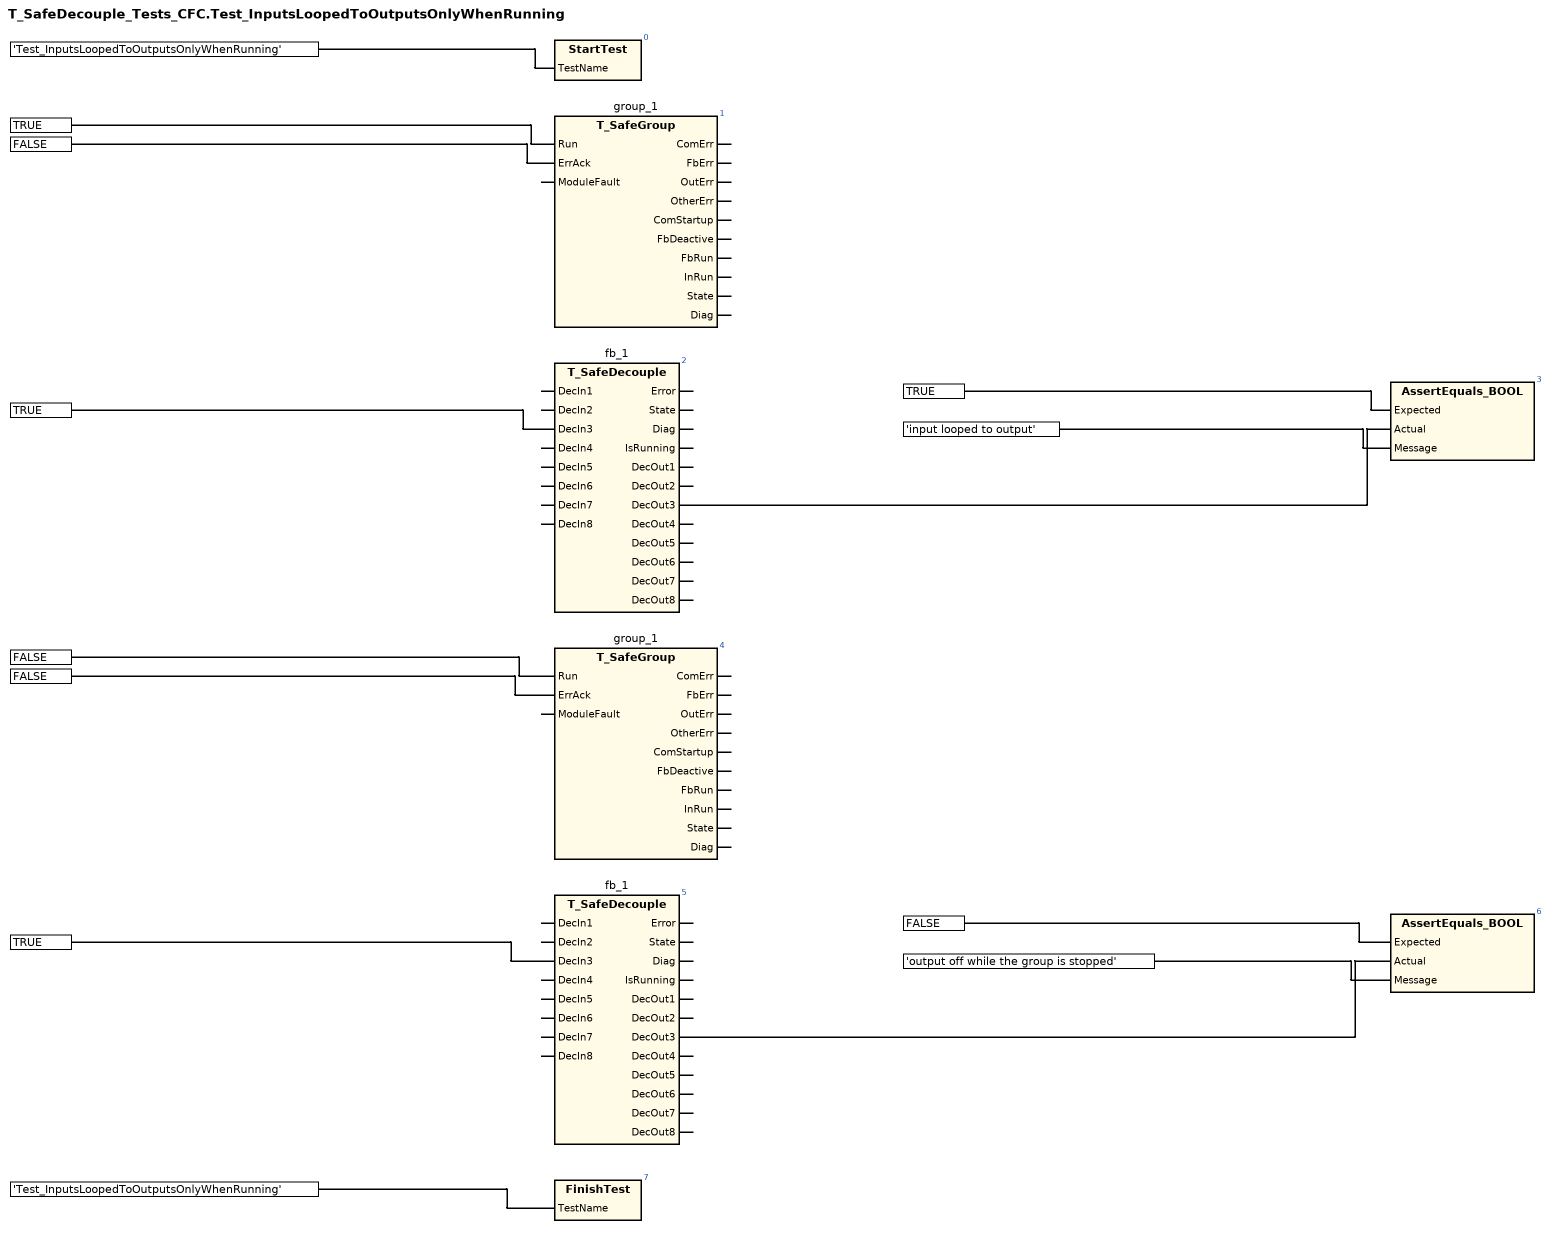
StartTest(TestName := 'Test_InputsLoopedToOutputsOnlyWhenRunning');
group_1(Run := TRUE, ErrAck := FALSE); // T_SafeGroup
fb_1(DecIn3 := TRUE); // T_SafeDecouple
AssertEquals_BOOL(Expected := TRUE, Actual := fb_1.DecOut3, Message := 'input looped to output');
group_1(Run := FALSE, ErrAck := FALSE); // T_SafeGroup
fb_1(DecIn3 := TRUE); // T_SafeDecouple
AssertEquals_BOOL(Expected := FALSE, Actual := fb_1.DecOut3, Message := 'output off while the group is stopped');
FinishTest(TestName := 'Test_InputsLoopedToOutputsOnlyWhenRunning');
END_METHOD

END_FUNCTION_BLOCK

// Tests/T_SafeOpMode_Tests_CFC
    // CFC twin of T_SafeOpMode_Tests: the same tests drawn as CFC diagrams, the way a TwinSAFE project is authored.
    FUNCTION_BLOCK T_SafeOpMode_Tests_CFC EXTENDS T_SafeCfcTestSuite
    VAR
    // Test_ExactlyOneInputSelectsOutput
    group_1 : T_SafeGroup;
    fb_1 : T_SafeOpMode(group := group_1);
    // Test_ConnectedRestartRequiresRestartSequence
    group_2 : T_SafeGroup;
    fb_2 : T_SafeOpMode(group := group_2);
    // Test_SlowModeChangeGivesDiscrepancyError
    group_3 : T_SafeGroup;
    fb_3 : T_SafeOpMode(group := group_3) := (Parameters := (DiscrepancyTime := T#100MS));
    t0_3 : TON;
    t1_3 : TON;
    trig1_3 : R_TRIG;
END_VAR

Test_ExactlyOneInputSelectsOutput();
Test_ConnectedRestartRequiresRestartSequence();
Test_SlowModeChangeGivesDiscrepancyError();

METHOD PRIVATE Test_ConnectedRestartRequiresRestartSequence
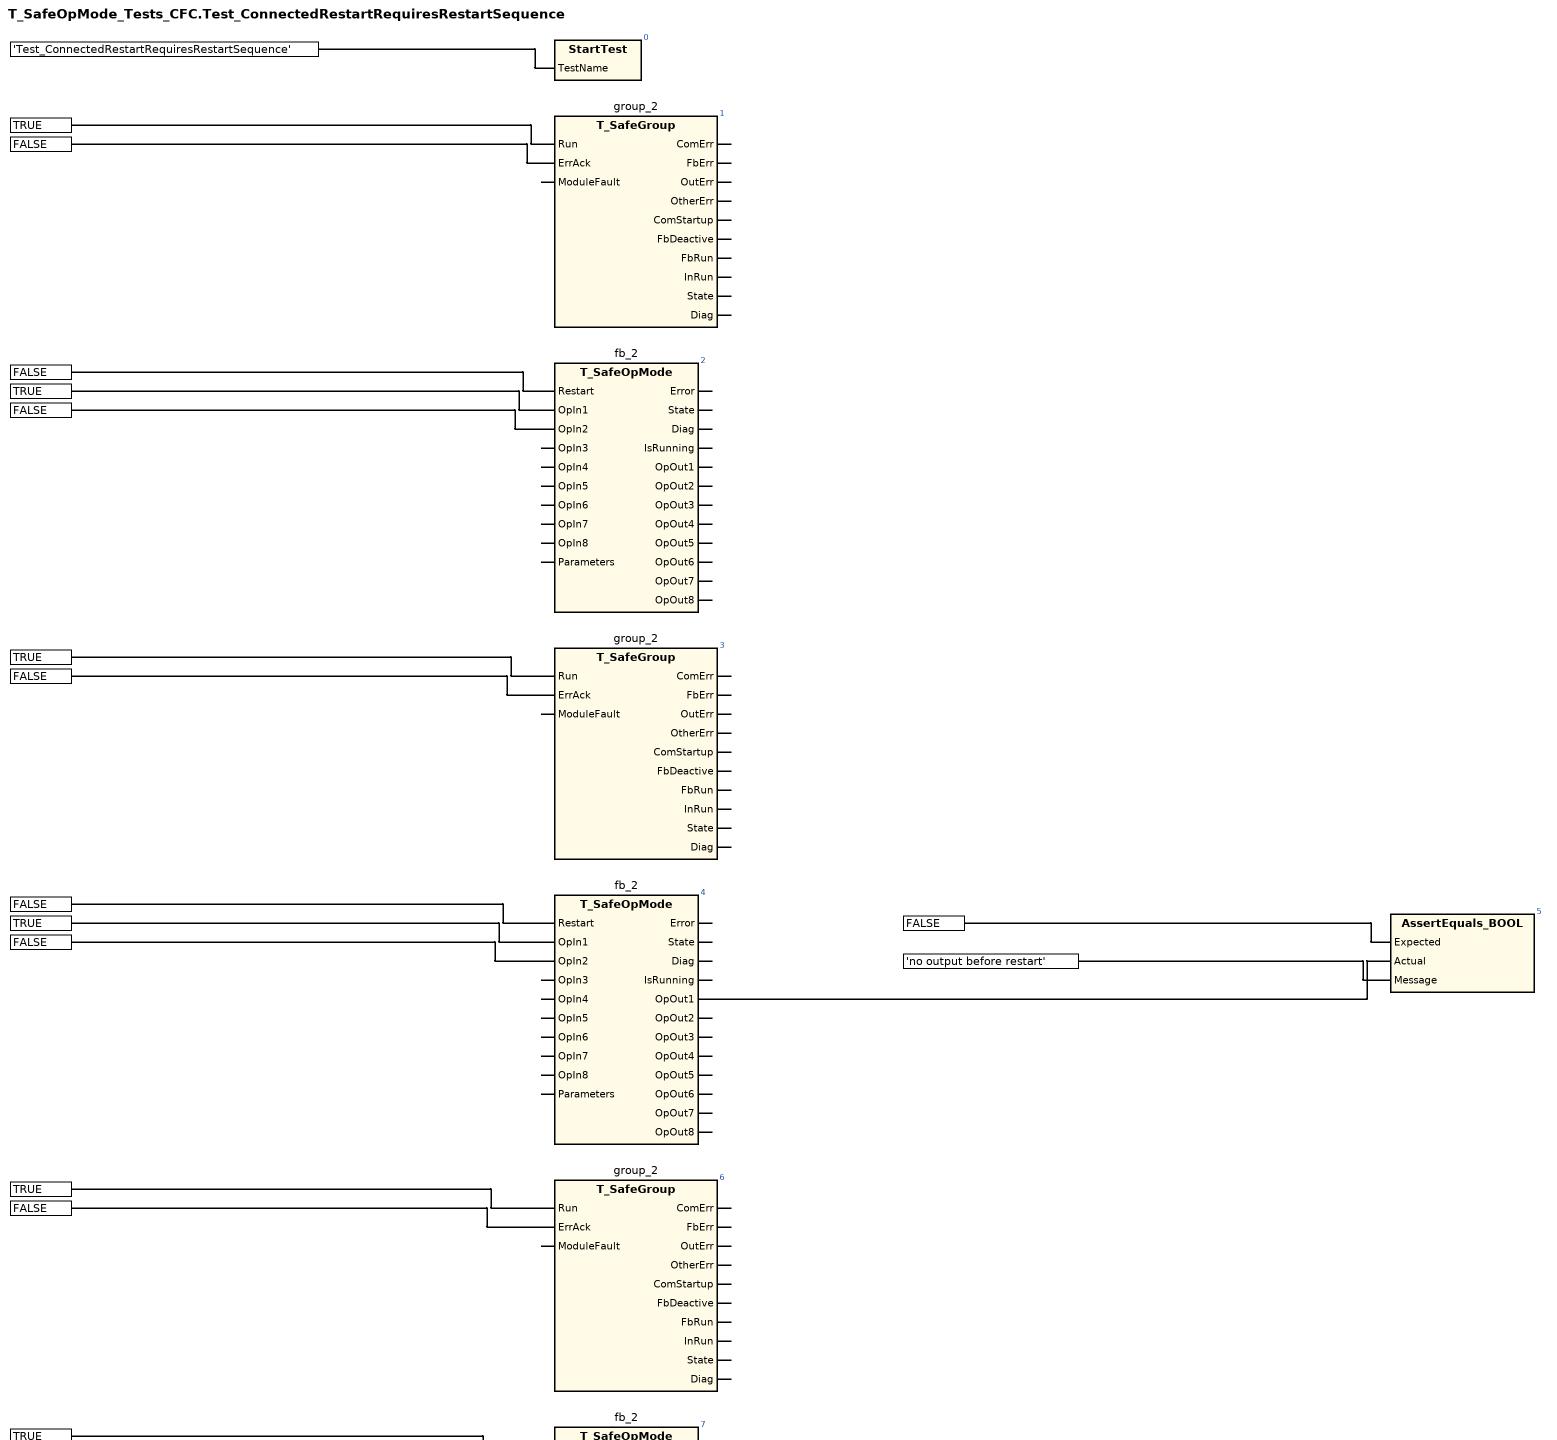
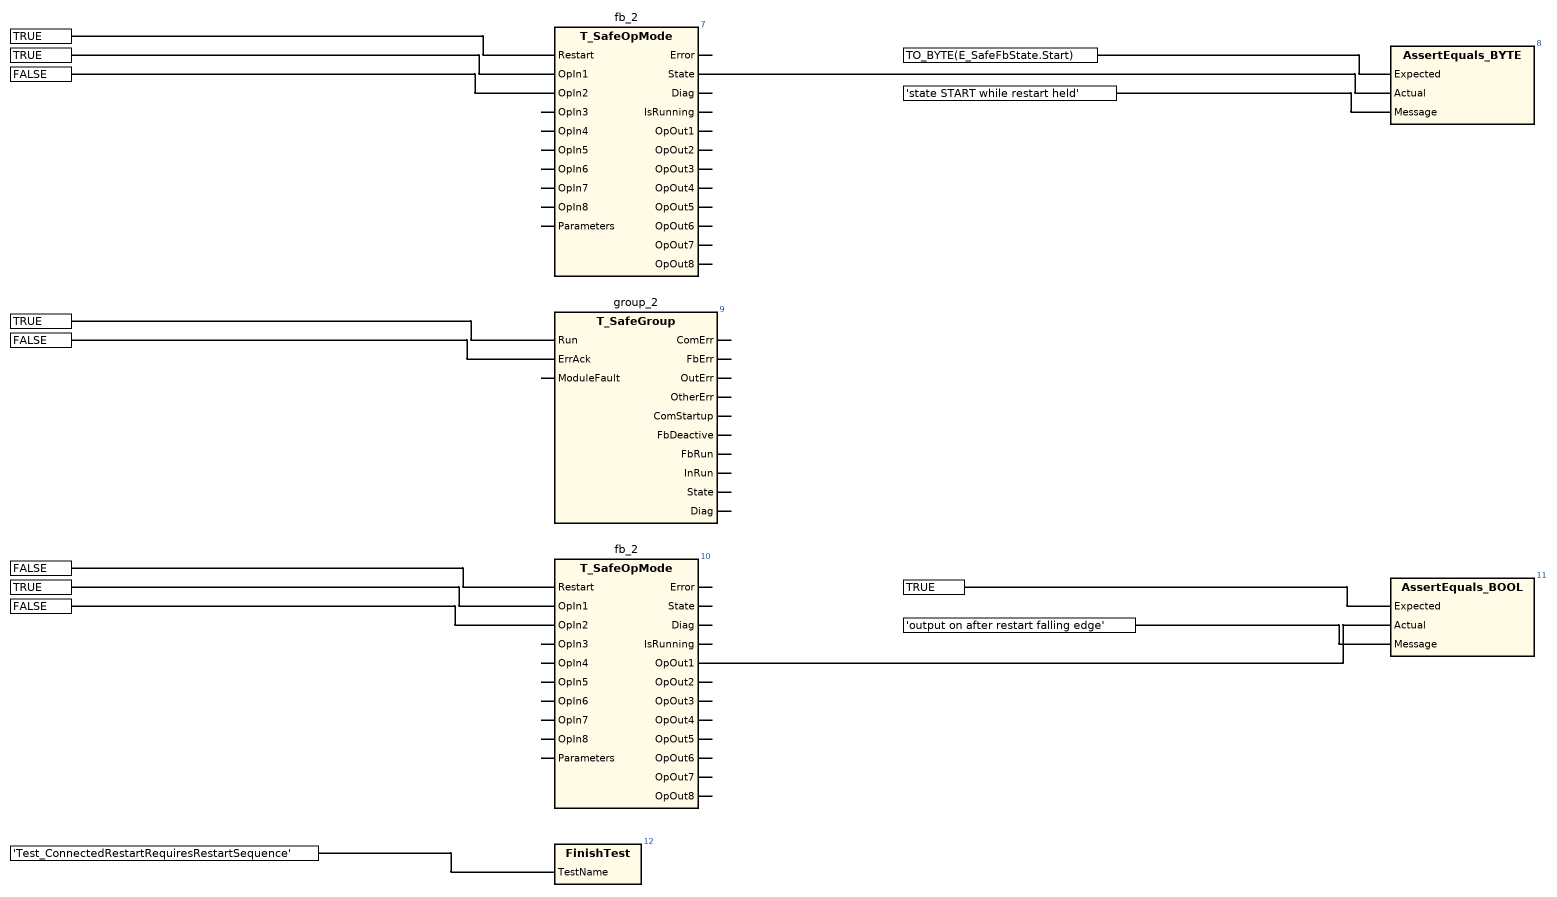
StartTest(TestName := 'Test_ConnectedRestartRequiresRestartSequence');
group_2(Run := TRUE, ErrAck := FALSE); // T_SafeGroup
fb_2(Restart := FALSE, OpIn1 := TRUE, OpIn2 := FALSE); // T_SafeOpMode
group_2(Run := TRUE, ErrAck := FALSE); // T_SafeGroup
fb_2(Restart := FALSE, OpIn1 := TRUE, OpIn2 := FALSE); // T_SafeOpMode
AssertEquals_BOOL(Expected := FALSE, Actual := fb_2.OpOut1, Message := 'no output before restart');
group_2(Run := TRUE, ErrAck := FALSE); // T_SafeGroup
fb_2(Restart := TRUE, OpIn1 := TRUE, OpIn2 := FALSE); // T_SafeOpMode
AssertEquals_BYTE(Expected := TO_BYTE(E_SafeFbState.Start), Actual := fb_2.State, Message := 'state START while restart held');
group_2(Run := TRUE, ErrAck := FALSE); // T_SafeGroup
fb_2(Restart := FALSE, OpIn1 := TRUE, OpIn2 := FALSE); // T_SafeOpMode
AssertEquals_BOOL(Expected := TRUE, Actual := fb_2.OpOut1, Message := 'output on after restart falling edge');
FinishTest(TestName := 'Test_ConnectedRestartRequiresRestartSequence');
END_METHOD

METHOD PRIVATE Test_ExactlyOneInputSelectsOutput
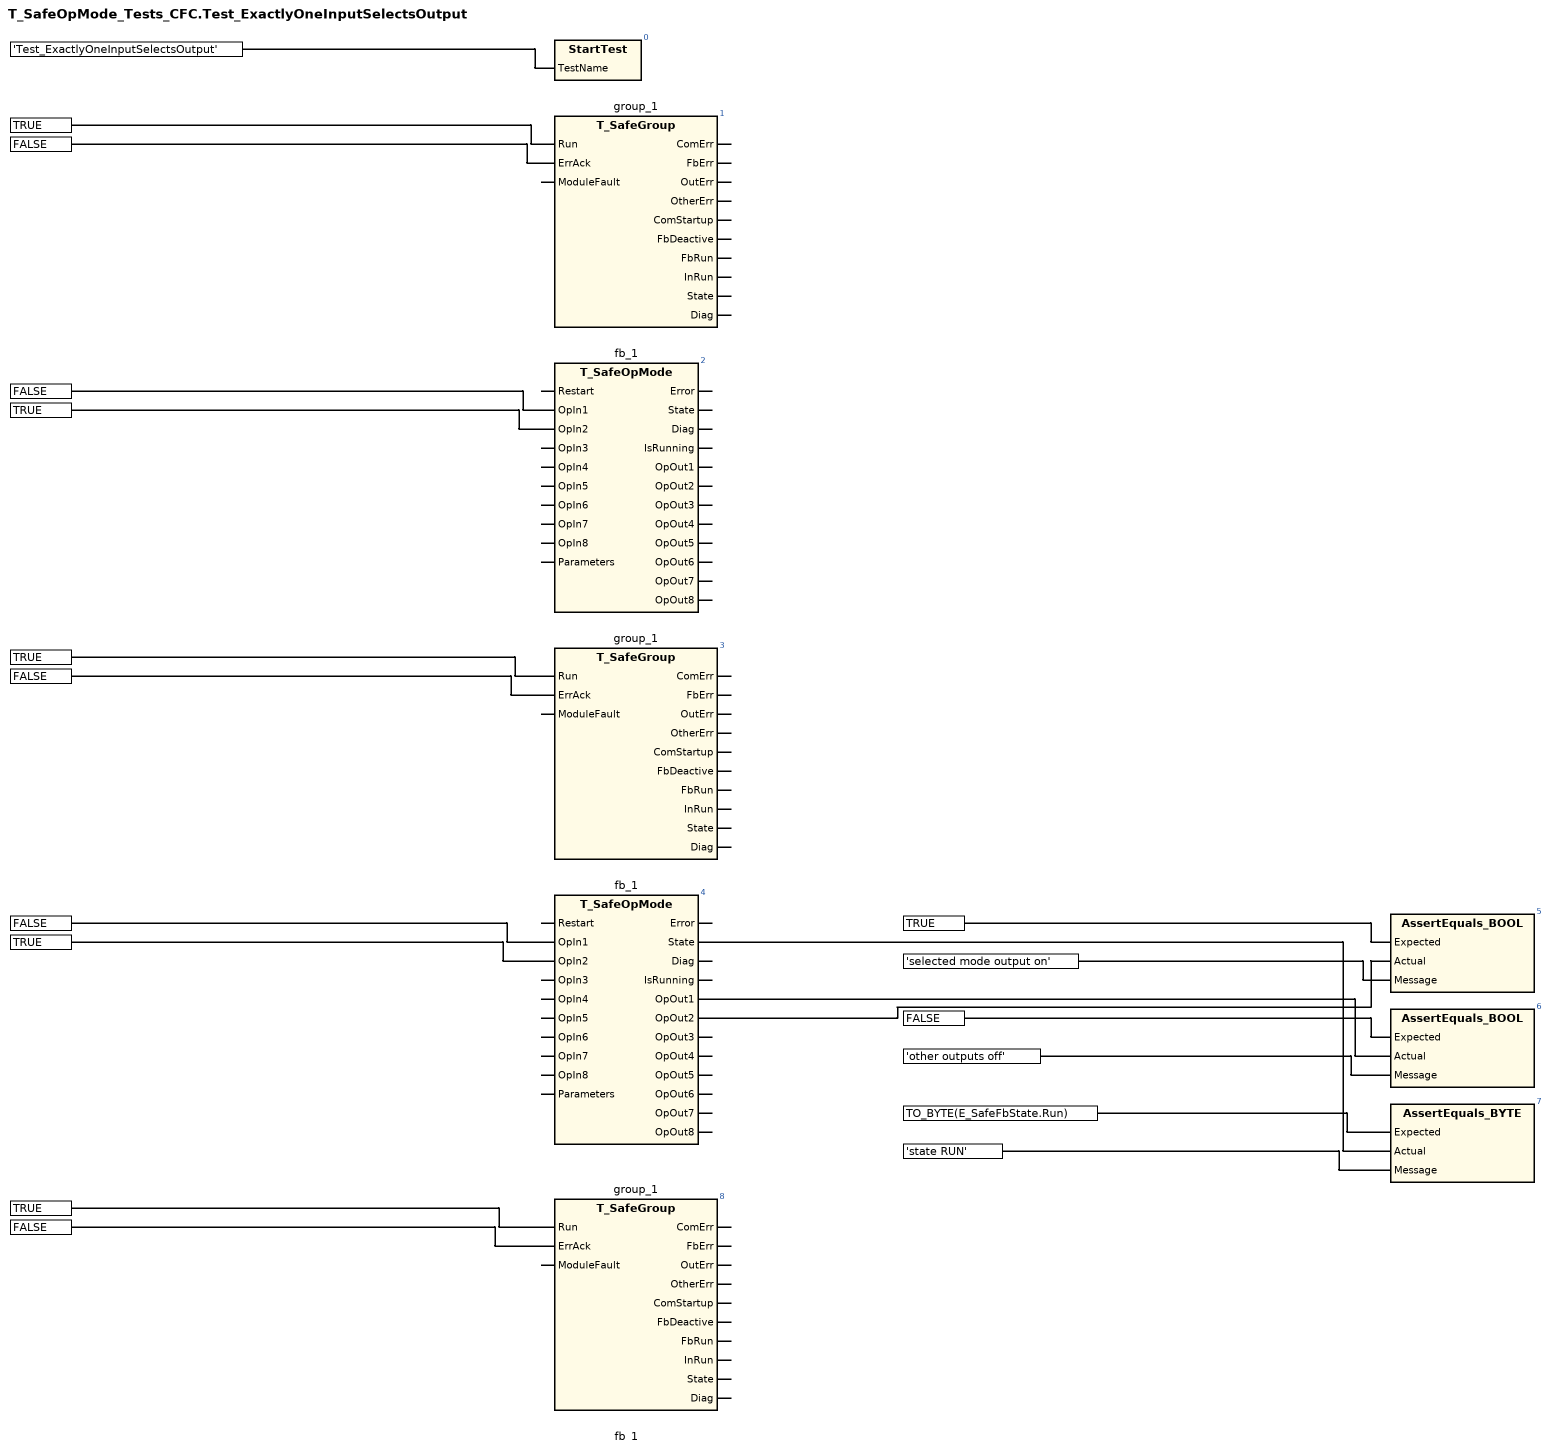
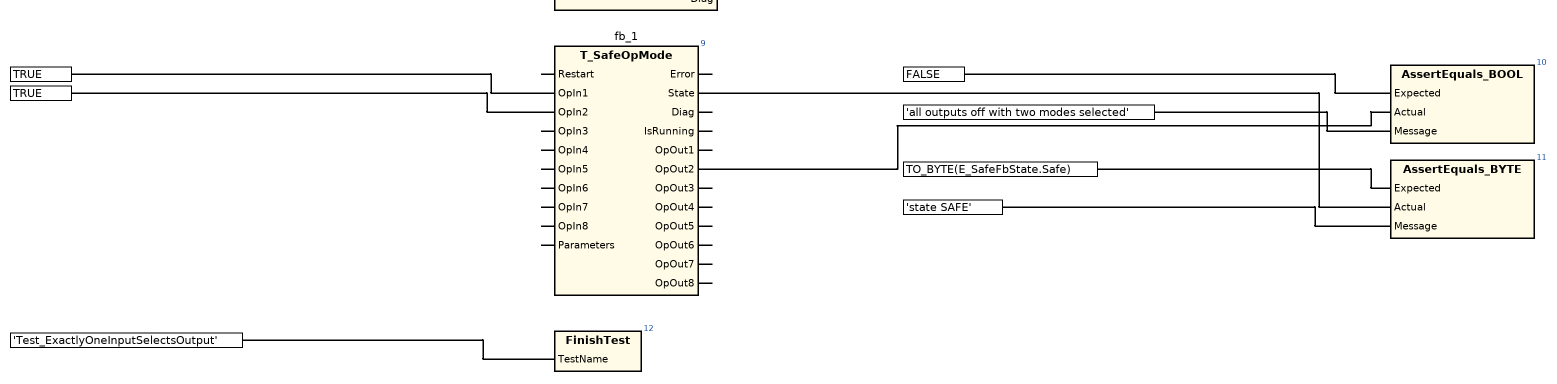
StartTest(TestName := 'Test_ExactlyOneInputSelectsOutput');
group_1(Run := TRUE, ErrAck := FALSE); // T_SafeGroup
fb_1(OpIn1 := FALSE, OpIn2 := TRUE); // T_SafeOpMode
group_1(Run := TRUE, ErrAck := FALSE); // T_SafeGroup
fb_1(OpIn1 := FALSE, OpIn2 := TRUE); // T_SafeOpMode
AssertEquals_BOOL(Expected := TRUE, Actual := fb_1.OpOut2, Message := 'selected mode output on');
AssertEquals_BOOL(Expected := FALSE, Actual := fb_1.OpOut1, Message := 'other outputs off');
AssertEquals_BYTE(Expected := TO_BYTE(E_SafeFbState.Run), Actual := fb_1.State, Message := 'state RUN');
group_1(Run := TRUE, ErrAck := FALSE); // T_SafeGroup
fb_1(OpIn1 := TRUE, OpIn2 := TRUE); // T_SafeOpMode
AssertEquals_BOOL(Expected := FALSE, Actual := fb_1.OpOut2, Message := 'all outputs off with two modes selected');
AssertEquals_BYTE(Expected := TO_BYTE(E_SafeFbState.Safe), Actual := fb_1.State, Message := 'state SAFE');
FinishTest(TestName := 'Test_ExactlyOneInputSelectsOutput');
END_METHOD

METHOD PRIVATE Test_SlowModeChangeGivesDiscrepancyError
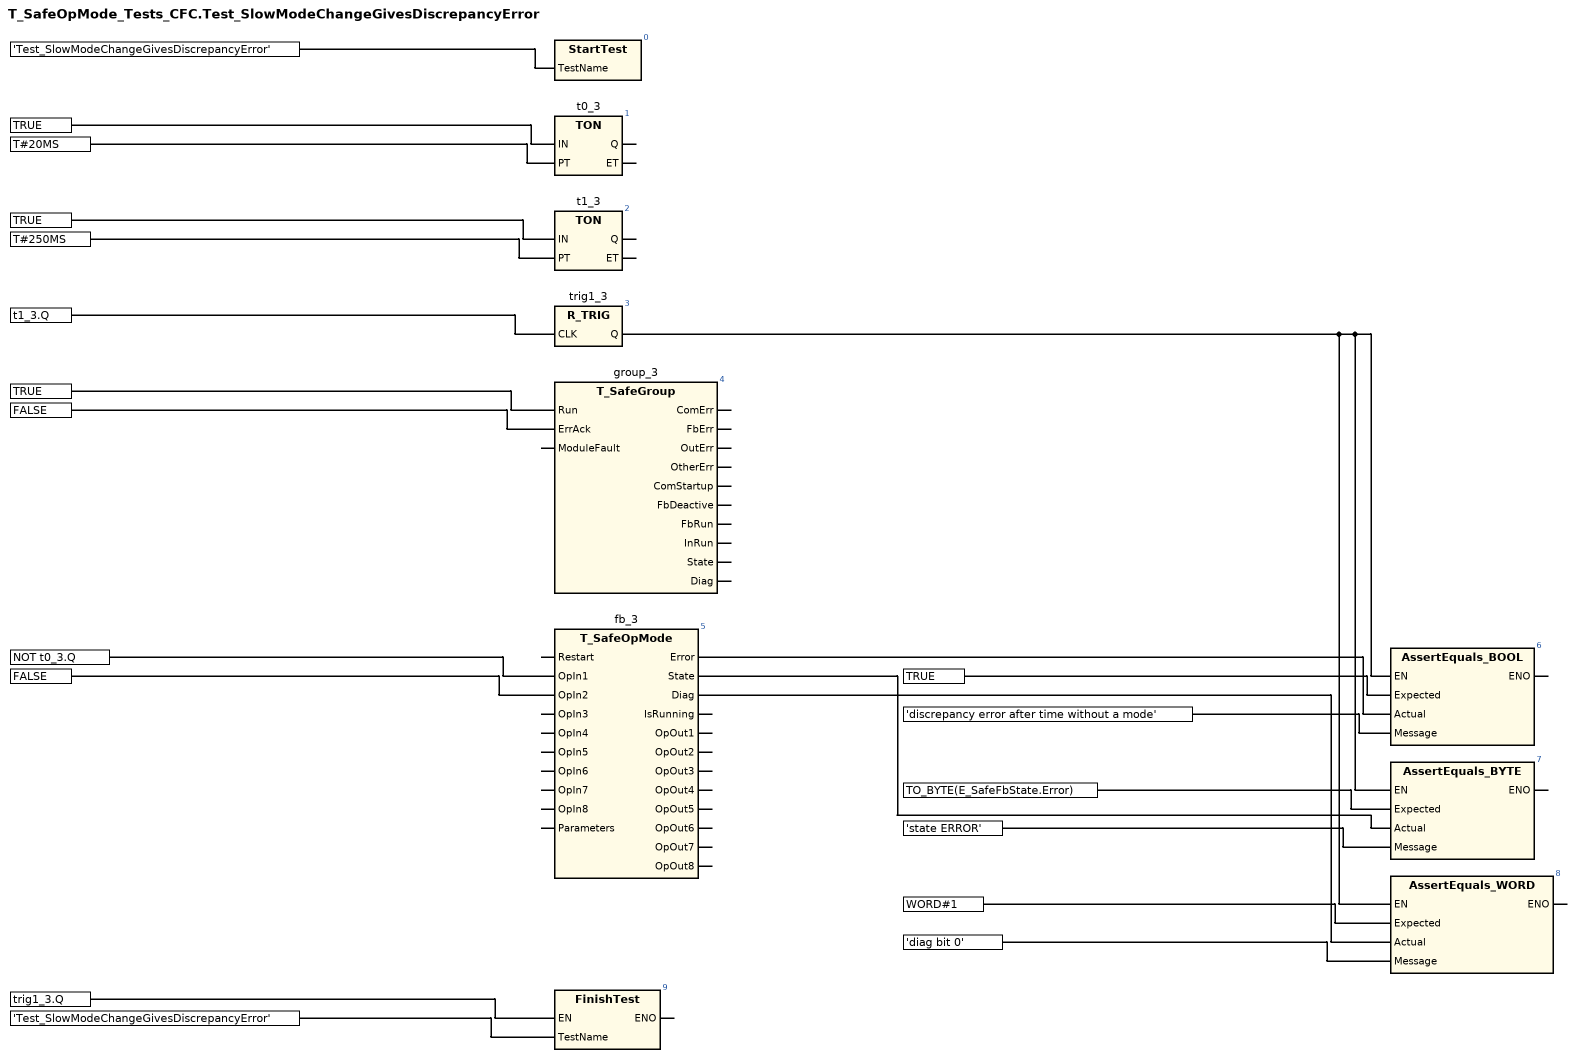
StartTest(TestName := 'Test_SlowModeChangeGivesDiscrepancyError');
t0_3(IN := TRUE, PT := T#20MS); // TON
t1_3(IN := TRUE, PT := T#250MS); // TON
trig1_3(CLK := t1_3.Q); // R_TRIG
group_3(Run := TRUE, ErrAck := FALSE); // T_SafeGroup
fb_3(OpIn1 := NOT t0_3.Q, OpIn2 := FALSE); // T_SafeOpMode
IF trig1_3.Q THEN AssertEquals_BOOL(Expected := TRUE, Actual := fb_3.Error, Message := 'discrepancy error after time without a mode'); END_IF
IF trig1_3.Q THEN AssertEquals_BYTE(Expected := TO_BYTE(E_SafeFbState.Error), Actual := fb_3.State, Message := 'state ERROR'); END_IF
IF trig1_3.Q THEN AssertEquals_WORD(Expected := WORD#1, Actual := fb_3.Diag, Message := 'diag bit 0'); END_IF
IF trig1_3.Q THEN FinishTest(TestName := 'Test_SlowModeChangeGivesDiscrepancyError'); END_IF
END_METHOD

END_FUNCTION_BLOCK

// Tests/T_SafeRs_Tests_CFC
    // CFC twin of T_SafeRs_Tests: the same tests drawn as CFC diagrams, the way a TwinSAFE project is authored.
    FUNCTION_BLOCK T_SafeRs_Tests_CFC EXTENDS T_SafeCfcTestSuite
    VAR
    // Test_ResetDominantLatch
    group_1 : T_SafeGroup;
    fb_1 : T_SafeRs(group := group_1);
END_VAR

Test_ResetDominantLatch();

METHOD PRIVATE Test_ResetDominantLatch
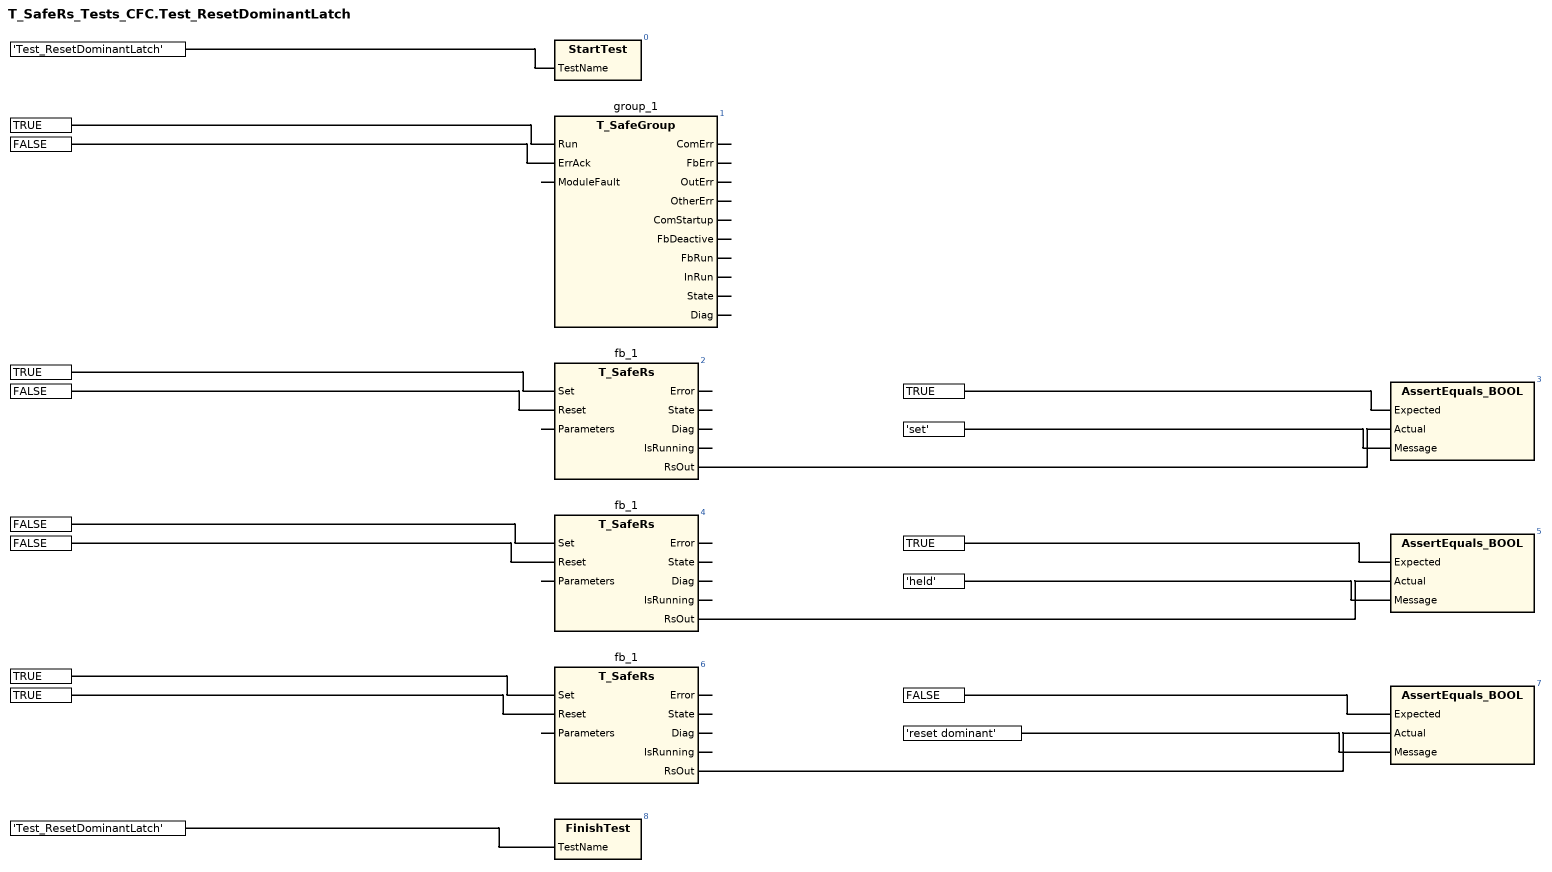
StartTest(TestName := 'Test_ResetDominantLatch');
group_1(Run := TRUE, ErrAck := FALSE); // T_SafeGroup
fb_1(Set := TRUE, Reset := FALSE); // T_SafeRs
AssertEquals_BOOL(Expected := TRUE, Actual := fb_1.RsOut, Message := 'set');
fb_1(Set := FALSE, Reset := FALSE); // T_SafeRs
AssertEquals_BOOL(Expected := TRUE, Actual := fb_1.RsOut, Message := 'held');
fb_1(Set := TRUE, Reset := TRUE); // T_SafeRs
AssertEquals_BOOL(Expected := FALSE, Actual := fb_1.RsOut, Message := 'reset dominant');
FinishTest(TestName := 'Test_ResetDominantLatch');
END_METHOD

END_FUNCTION_BLOCK

// Tests/T_SafeSr_Tests_CFC
    // CFC twin of T_SafeSr_Tests: the same tests drawn as CFC diagrams, the way a TwinSAFE project is authored.
    FUNCTION_BLOCK T_SafeSr_Tests_CFC EXTENDS T_SafeCfcTestSuite
    VAR
    // Test_SetDominantLatch
    group_1 : T_SafeGroup;
    fb_1 : T_SafeSr(group := group_1);
END_VAR

Test_SetDominantLatch();

METHOD PRIVATE Test_SetDominantLatch
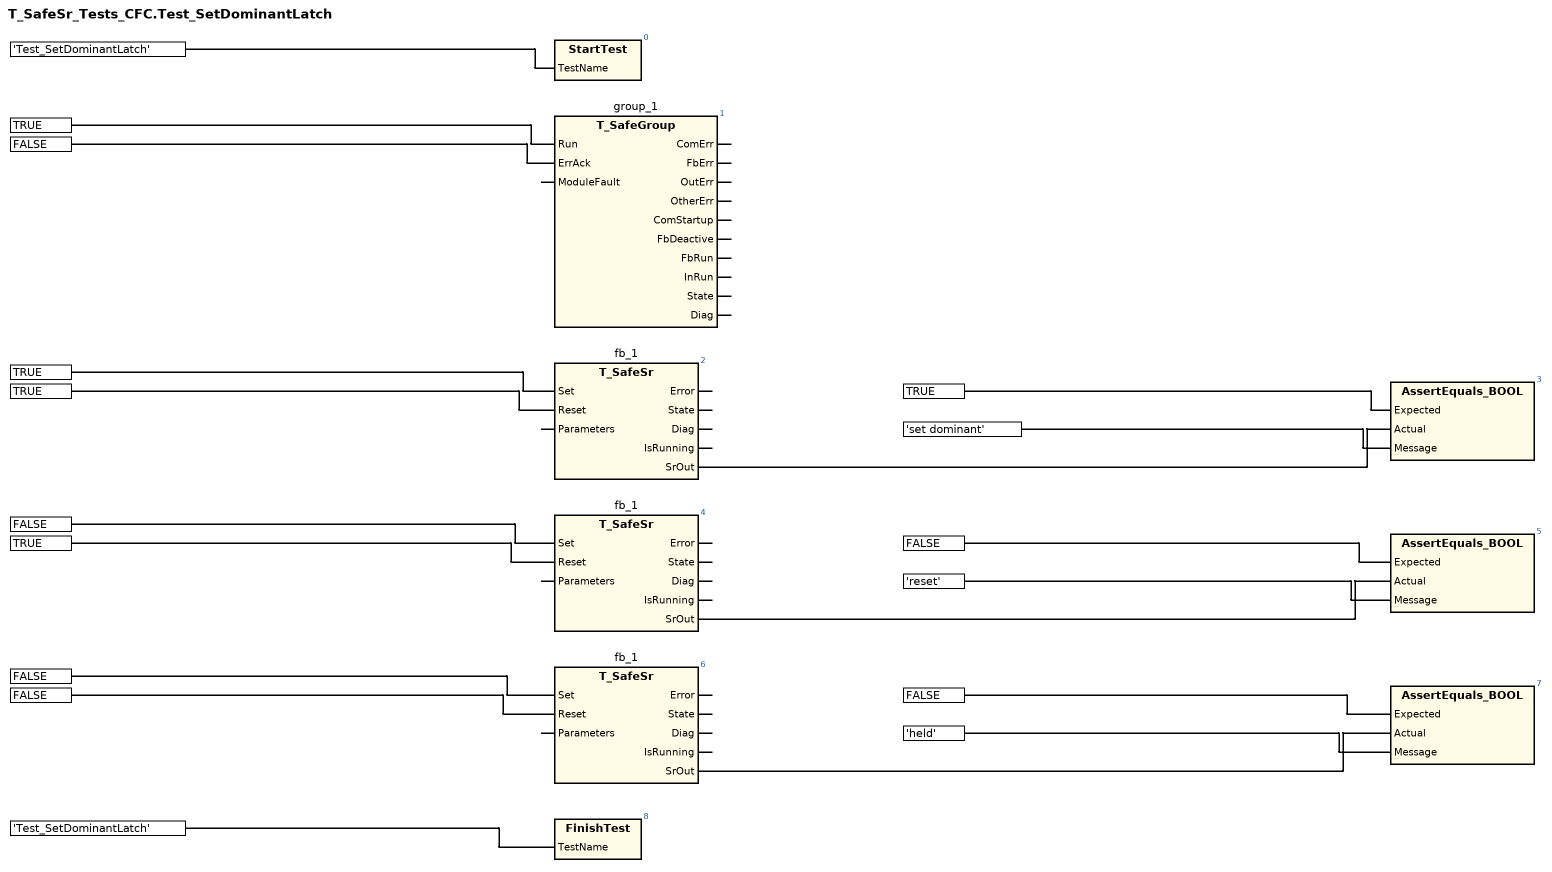
StartTest(TestName := 'Test_SetDominantLatch');
group_1(Run := TRUE, ErrAck := FALSE); // T_SafeGroup
fb_1(Set := TRUE, Reset := TRUE); // T_SafeSr
AssertEquals_BOOL(Expected := TRUE, Actual := fb_1.SrOut, Message := 'set dominant');
fb_1(Set := FALSE, Reset := TRUE); // T_SafeSr
AssertEquals_BOOL(Expected := FALSE, Actual := fb_1.SrOut, Message := 'reset');
fb_1(Set := FALSE, Reset := FALSE); // T_SafeSr
AssertEquals_BOOL(Expected := FALSE, Actual := fb_1.SrOut, Message := 'held');
FinishTest(TestName := 'Test_SetDominantLatch');
END_METHOD

END_FUNCTION_BLOCK

// Tests/T_SafeTon_Tests_CFC
    // CFC twin of T_SafeTon_Tests: the same tests drawn as CFC diagrams, the way a TwinSAFE project is authored.
    FUNCTION_BLOCK T_SafeTon_Tests_CFC EXTENDS T_SafeCfcTestSuite
    VAR
    // Test_OutputDelayedOn
    group_1 : T_SafeGroup;
    fb_1 : T_SafeTon(group := group_1) := (Parameters := (DelayTime := T#100MS));
    trigStart_1 : R_TRIG;
    t1_1 : TON;
    trig1_1 : R_TRIG;
END_VAR

Test_OutputDelayedOn();

METHOD PRIVATE Test_OutputDelayedOn
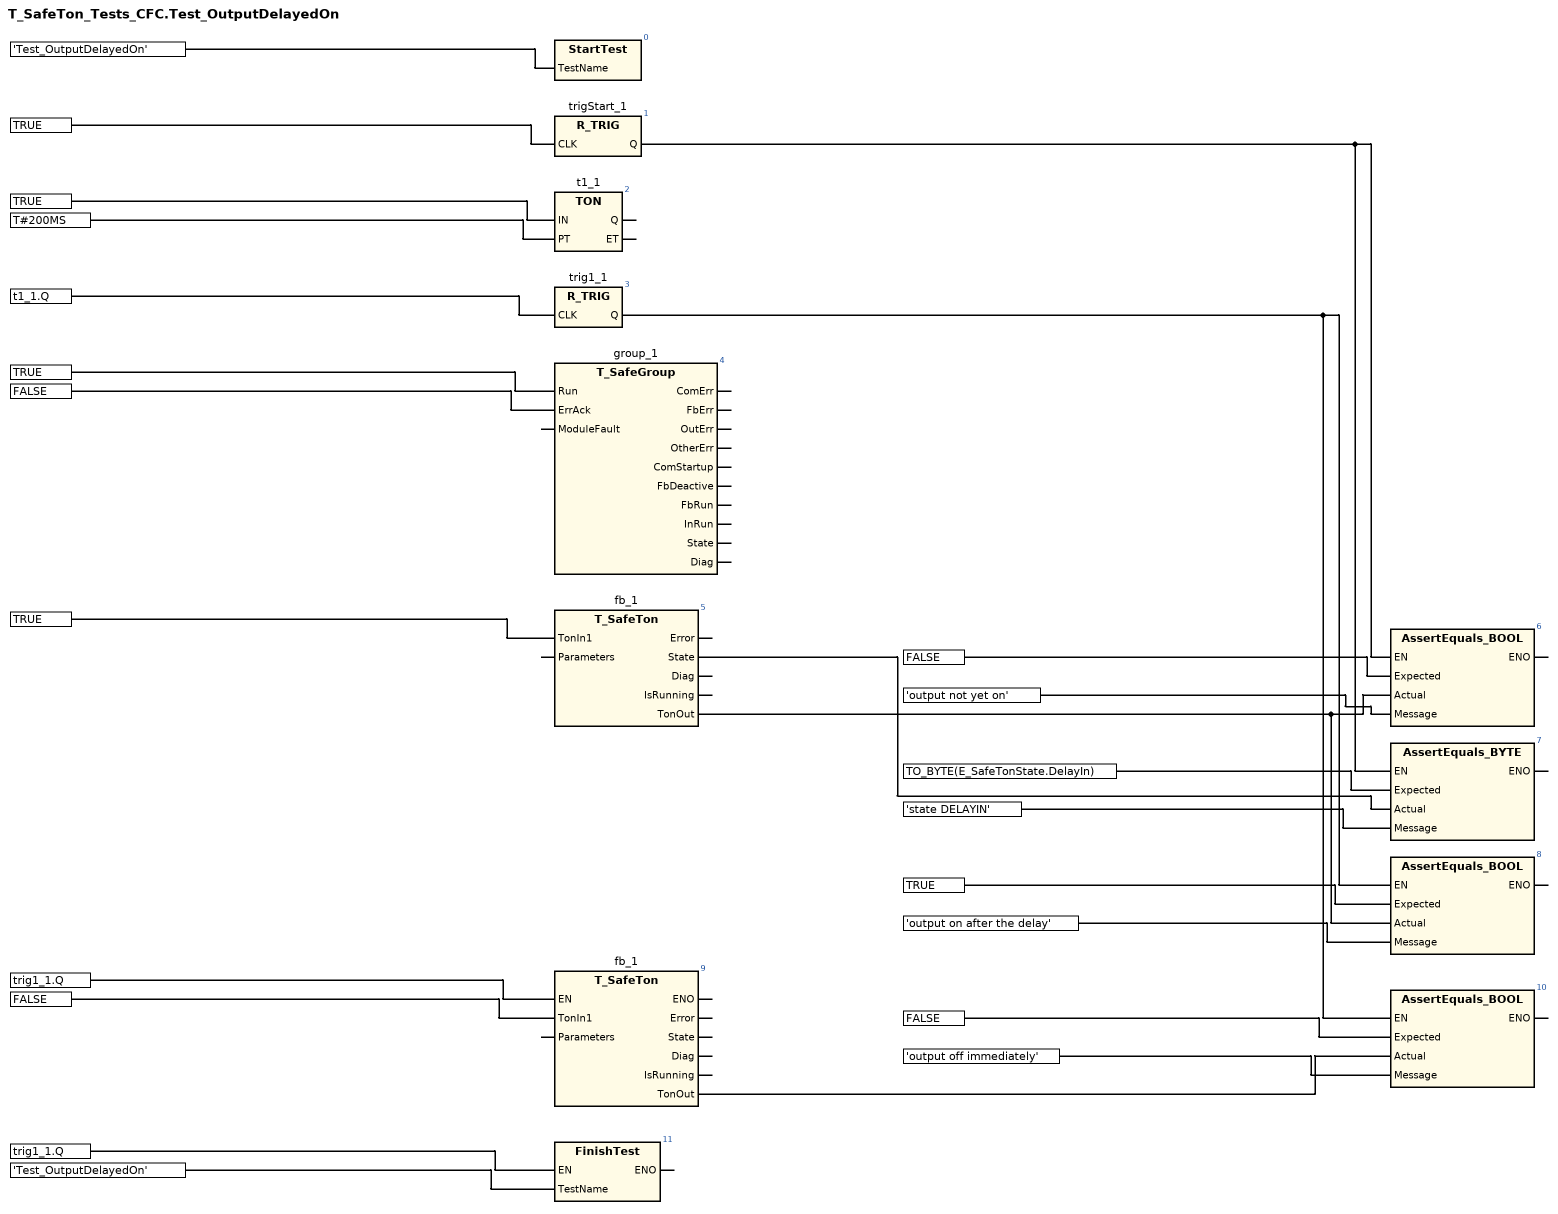
StartTest(TestName := 'Test_OutputDelayedOn');
trigStart_1(CLK := TRUE); // R_TRIG
t1_1(IN := TRUE, PT := T#200MS); // TON
trig1_1(CLK := t1_1.Q); // R_TRIG
group_1(Run := TRUE, ErrAck := FALSE); // T_SafeGroup
fb_1(TonIn1 := TRUE); // T_SafeTon
IF trigStart_1.Q THEN AssertEquals_BOOL(Expected := FALSE, Actual := fb_1.TonOut, Message := 'output not yet on'); END_IF
IF trigStart_1.Q THEN AssertEquals_BYTE(Expected := TO_BYTE(E_SafeTonState.DelayIn), Actual := fb_1.State, Message := 'state DELAYIN'); END_IF
IF trig1_1.Q THEN AssertEquals_BOOL(Expected := TRUE, Actual := fb_1.TonOut, Message := 'output on after the delay'); END_IF
IF trig1_1.Q THEN
    fb_1(TonIn1 := FALSE); // T_SafeTon
END_IF
IF trig1_1.Q THEN AssertEquals_BOOL(Expected := FALSE, Actual := fb_1.TonOut, Message := 'output off immediately'); END_IF
IF trig1_1.Q THEN FinishTest(TestName := 'Test_OutputDelayedOn'); END_IF
END_METHOD

END_FUNCTION_BLOCK

// Tests/T_SafeTof_Tests_CFC
    // CFC twin of T_SafeTof_Tests: the same tests drawn as CFC diagrams, the way a TwinSAFE project is authored.
    FUNCTION_BLOCK T_SafeTof_Tests_CFC EXTENDS T_SafeCfcTestSuite
    VAR
    // Test_OutputDelayedOff
    group_1 : T_SafeGroup;
    fb_1 : T_SafeTof(group := group_1) := (Parameters := (DelayTime := T#100MS));
    trigStart_1 : R_TRIG;
    t0_1 : TON;
    t1_1 : TON;
    trig0_1 : R_TRIG;
    trig1_1 : R_TRIG;
END_VAR

Test_OutputDelayedOff();

METHOD PRIVATE Test_OutputDelayedOff
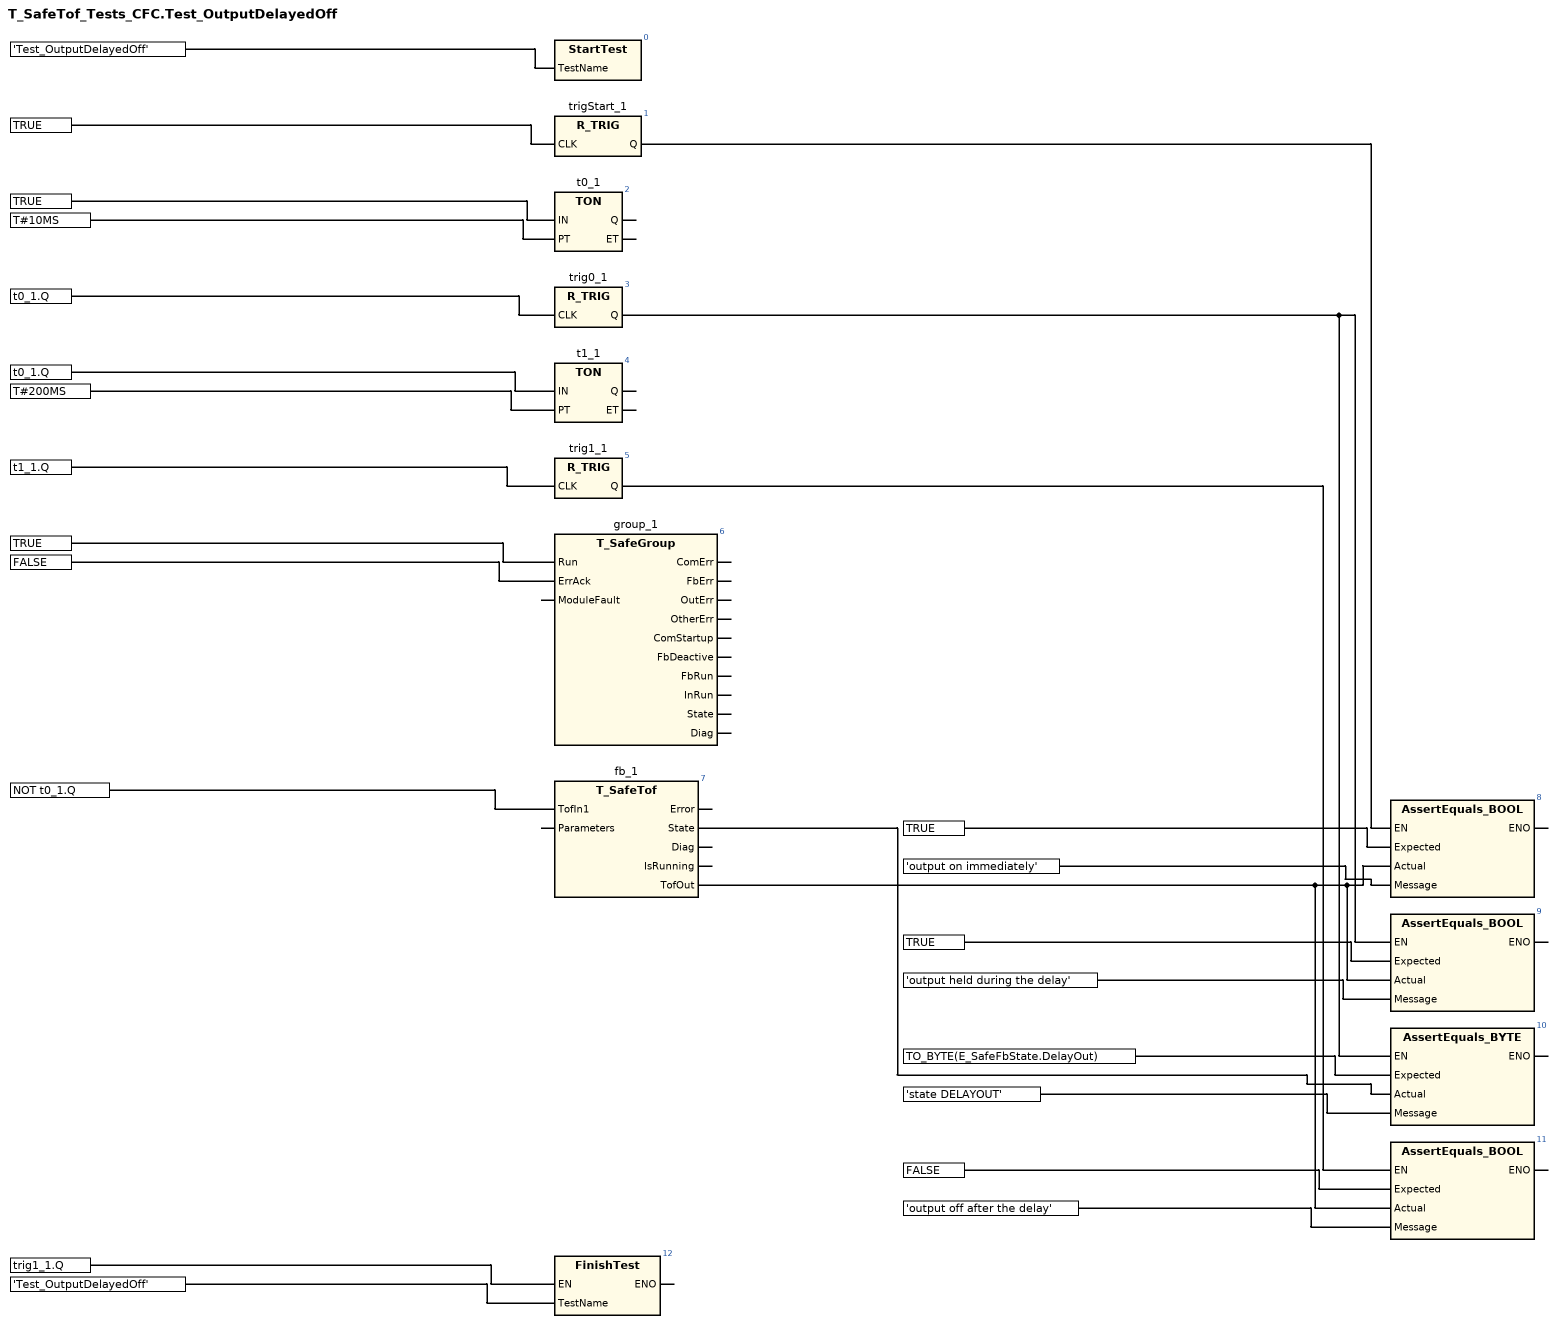
StartTest(TestName := 'Test_OutputDelayedOff');
trigStart_1(CLK := TRUE); // R_TRIG
t0_1(IN := TRUE, PT := T#10MS); // TON
trig0_1(CLK := t0_1.Q); // R_TRIG
t1_1(IN := t0_1.Q, PT := T#200MS); // TON
trig1_1(CLK := t1_1.Q); // R_TRIG
group_1(Run := TRUE, ErrAck := FALSE); // T_SafeGroup
fb_1(TofIn1 := NOT t0_1.Q); // T_SafeTof
IF trigStart_1.Q THEN AssertEquals_BOOL(Expected := TRUE, Actual := fb_1.TofOut, Message := 'output on immediately'); END_IF
IF trig0_1.Q THEN AssertEquals_BOOL(Expected := TRUE, Actual := fb_1.TofOut, Message := 'output held during the delay'); END_IF
IF trig0_1.Q THEN AssertEquals_BYTE(Expected := TO_BYTE(E_SafeFbState.DelayOut), Actual := fb_1.State, Message := 'state DELAYOUT'); END_IF
IF trig1_1.Q THEN AssertEquals_BOOL(Expected := FALSE, Actual := fb_1.TofOut, Message := 'output off after the delay'); END_IF
IF trig1_1.Q THEN FinishTest(TestName := 'Test_OutputDelayedOff'); END_IF
END_METHOD

END_FUNCTION_BLOCK

// Tests/T_SafeEdm_Tests_CFC
    // CFC twin of T_SafeEdm_Tests: the same tests drawn as CFC diagrams, the way a TwinSAFE project is authored.
    FUNCTION_BLOCK T_SafeEdm_Tests_CFC EXTENDS T_SafeCfcTestSuite
    VAR
    // Test_SwitchOnTimeoutGivesError
    group_1 : T_SafeGroup;
    fb_1 : T_SafeEdm(group := group_1) := (Parameters := (SwitchOnTime := T#100MS));
    t1_1 : TON;
    trig1_1 : R_TRIG;
    // Test_NoErrorWhenFeedbackFollows
    group_2 : T_SafeGroup;
    fb_2 : T_SafeEdm(group := group_2) := (Parameters := (SwitchOnTime := T#100MS, SwitchOffTime := T#100MS));
    t1_2 : TON;
    t2_2 : TON;
    trig1_2 : R_TRIG;
    trig2_2 : R_TRIG;
END_VAR

Test_SwitchOnTimeoutGivesError();
Test_NoErrorWhenFeedbackFollows();

METHOD PRIVATE Test_NoErrorWhenFeedbackFollows
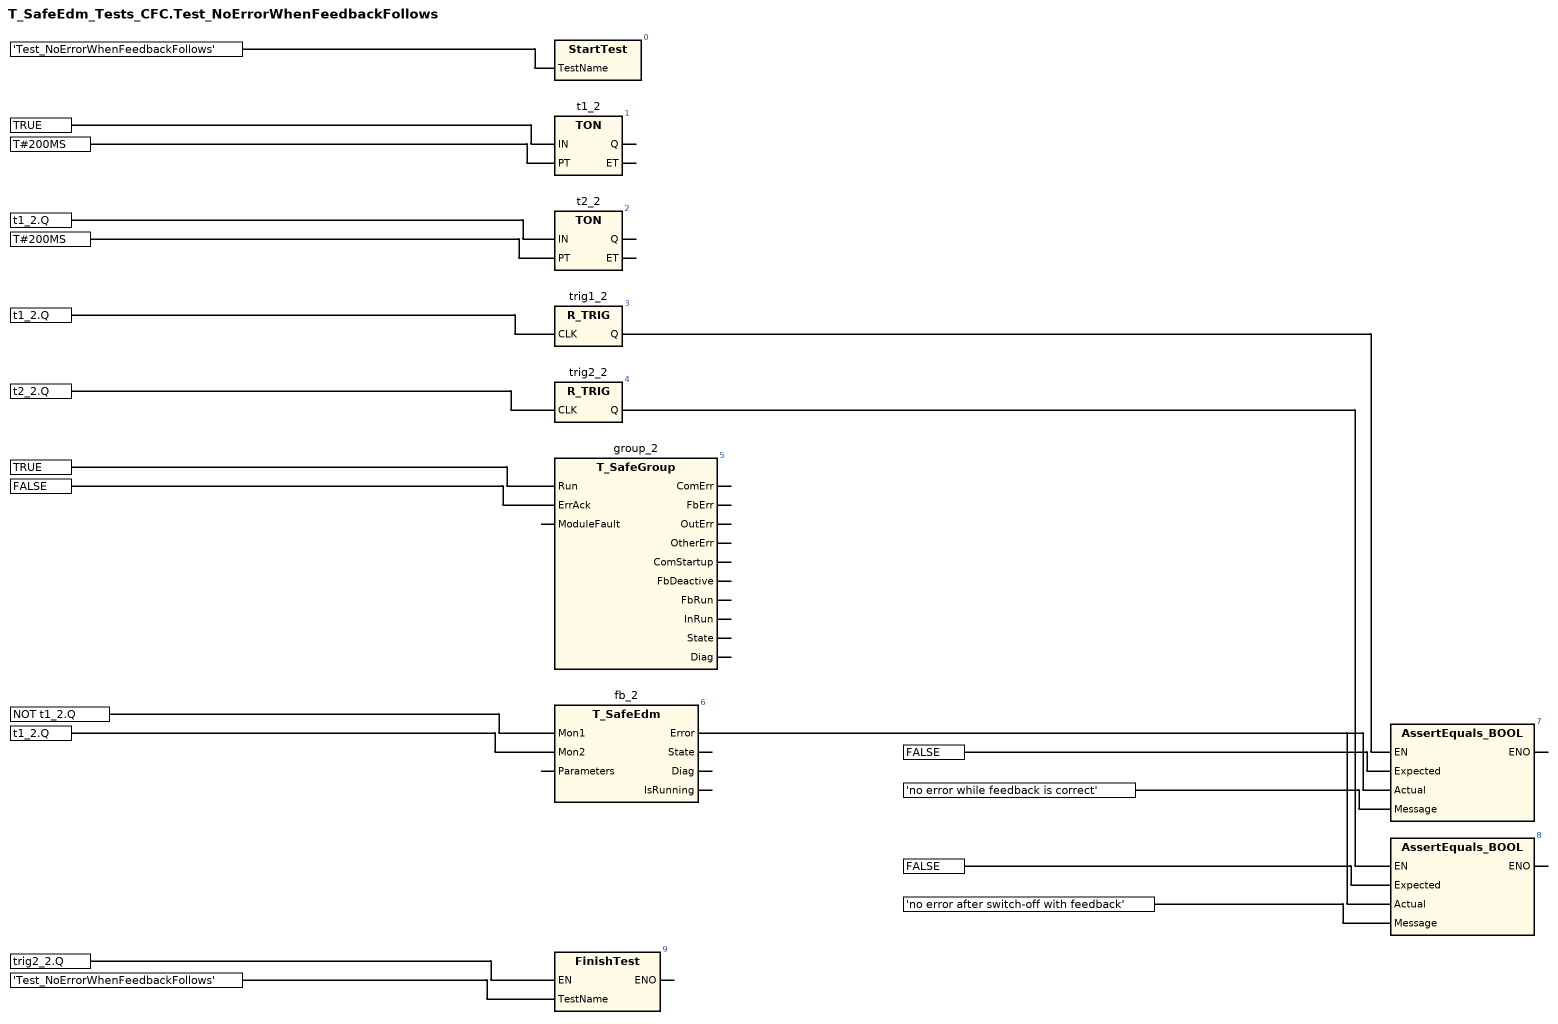
StartTest(TestName := 'Test_NoErrorWhenFeedbackFollows');
t1_2(IN := TRUE, PT := T#200MS); // TON
t2_2(IN := t1_2.Q, PT := T#200MS); // TON
trig1_2(CLK := t1_2.Q); // R_TRIG
trig2_2(CLK := t2_2.Q); // R_TRIG
group_2(Run := TRUE, ErrAck := FALSE); // T_SafeGroup
fb_2(Mon1 := NOT t1_2.Q, Mon2 := t1_2.Q); // T_SafeEdm
IF trig1_2.Q THEN AssertEquals_BOOL(Expected := FALSE, Actual := fb_2.Error, Message := 'no error while feedback is correct'); END_IF
IF trig2_2.Q THEN AssertEquals_BOOL(Expected := FALSE, Actual := fb_2.Error, Message := 'no error after switch-off with feedback'); END_IF
IF trig2_2.Q THEN FinishTest(TestName := 'Test_NoErrorWhenFeedbackFollows'); END_IF
END_METHOD

METHOD PRIVATE Test_SwitchOnTimeoutGivesError
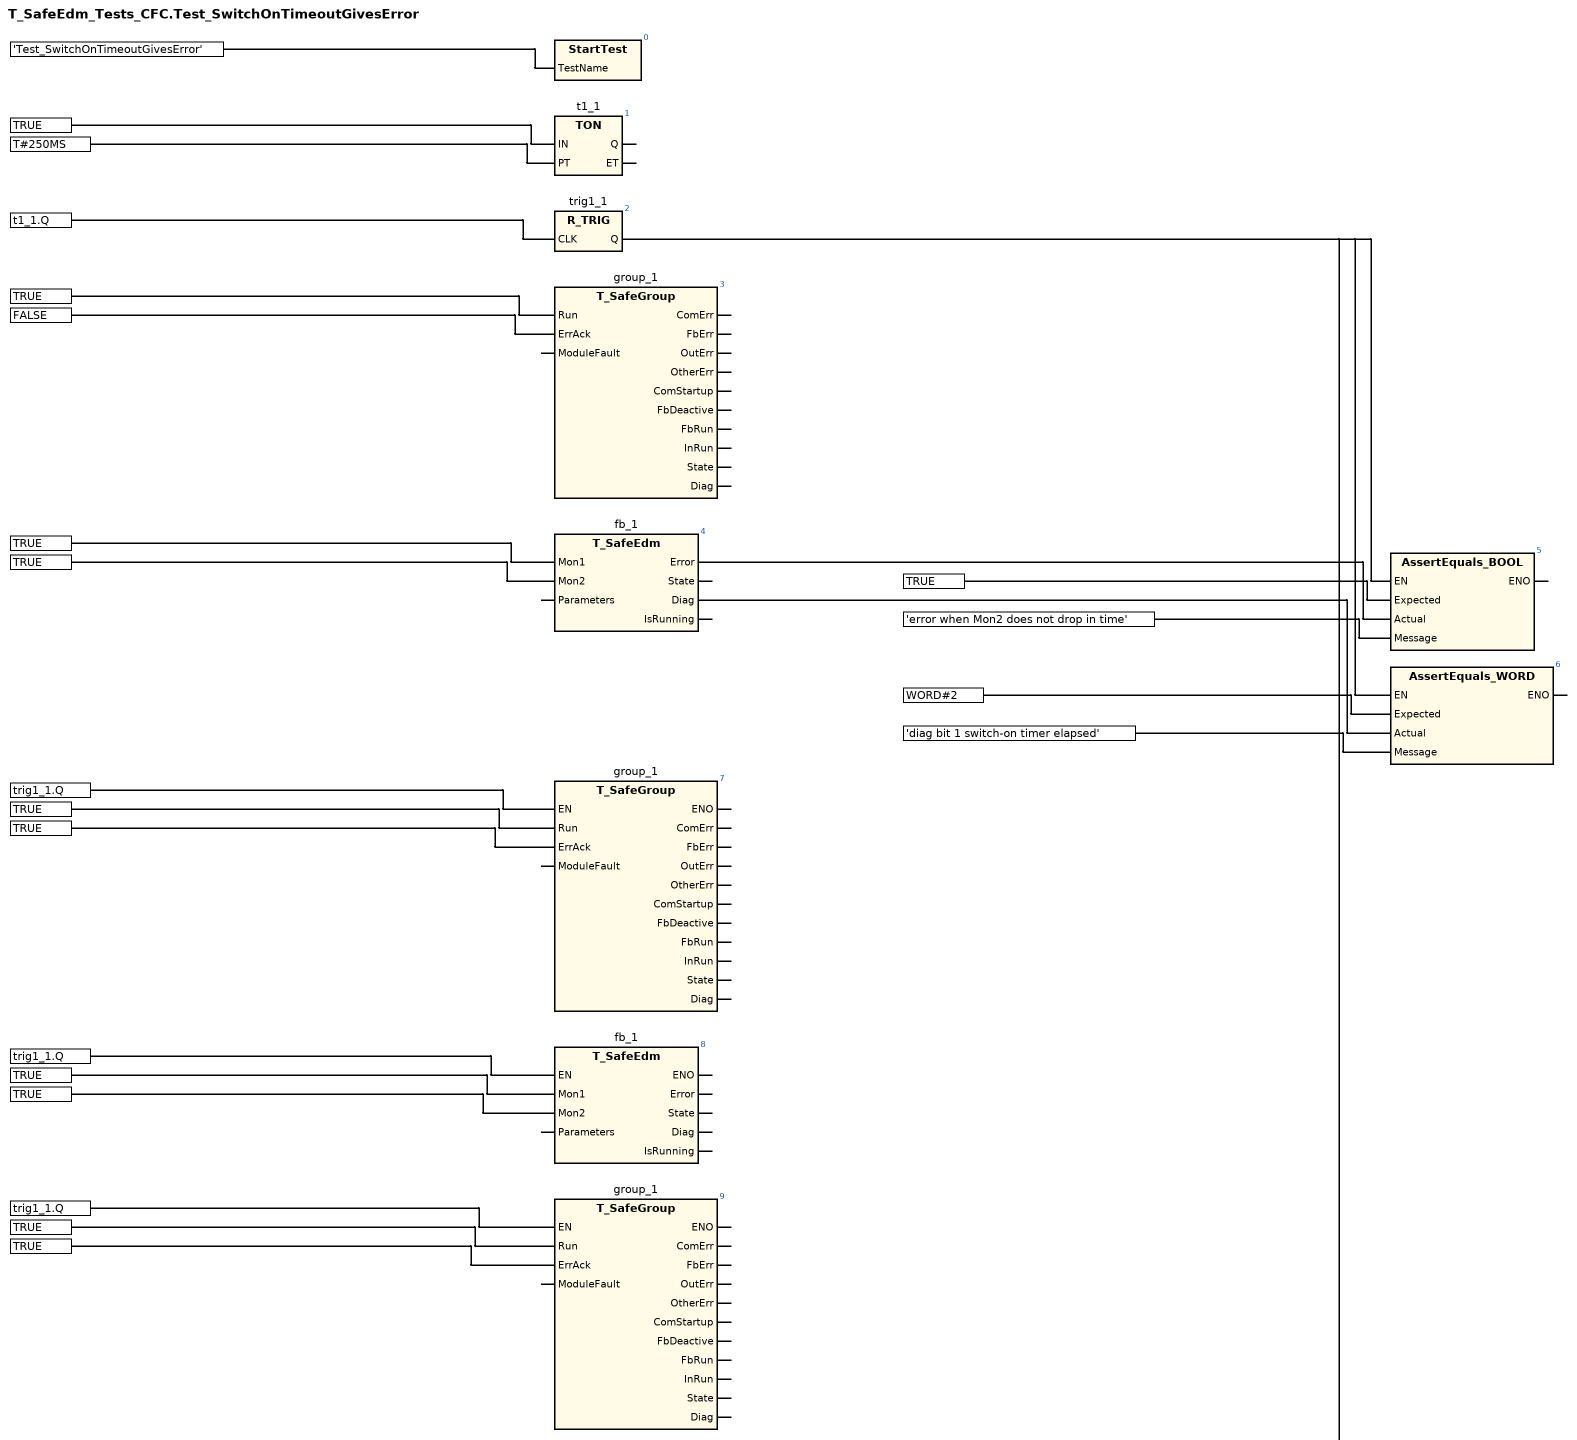
